The real Test Case computes reservations; the real Orchestrator decides and publishes its diagnostic.
A collection double supplies one fixed child view. Only the concurrent Suite allowance is held by
the fixture, without running a Suite. Request-entry observations are inherited from the thin child adapter.
The fault is injected by early FreeReservedEvents on a started child, not by corrupting indices or interfaces.
This tests the missing-reservation invariant; hard Event Buffer Reset mechanics are not reproduced.
Three later helper calls must retain Error without another diagnostic or unexpected dispatch.
Expected diagnostics stay in local capture. The surrounding Assertions use the normal selftest publisher.
The real subject binds only local storage; expected findings remain in that storage.
Checking Assertions retain the outer selftest publisher. Each run reinitializes the subject.
</description>
*)
{endregion}
FUNCTION_BLOCK Test_ActiveReservationLoss EXTENDS TestCaseBase
VAR
    FSubject : EventBuffer;
    FEvents : ARRAY[1..BufferLength] OF ST_Event;
    FFifo : ST_FifoStatus;
    FBufferStatus : ST_EventBufferStatus;
    FPerformed : BOOL;
    FChecked : BOOL;
    FSubjectParent : I_TestSuite;
    FChild : ReservationChildProbe;
    FOrchestrator : OrchestratorProbe;
    FCollection : OrchestrationCollectionDouble;
    FChildren : ARRAY[1..1] OF I_Orchestratable;
    FOwnerReserved : UINT;
    FStep : INT;
    FObservationCalls : UINT;
    FPrecondition : AssertTrue;
    FPreconditionMatches : BOOL;
    FFailureDetection : AssertTrue;
    FFailureDetectionMatches : BOOL;
    FStateAndCounts : AssertTrue;
    FStateAndCountsMatches : BOOL;
    FHeldError : AssertTrue;
    FHeldErrorMatches : BOOL;
    FSingleDiagnostic : AssertTrue;
    FSingleDiagnosticMatches : BOOL;
    FRequestBoundary : AssertTrue;
    FRequestBoundaryMatches : BOOL;
    FAccounting : AssertTrue;
    FAccountingMatches : BOOL;
    FCaptureIntegrity : AssertTrue;
    FCaptureIntegrityMatches : BOOL;
END_VAR
VAR CONSTANT
    ChildExecutionBudget : UINT := 11;
    ConfigureExecution : INT := 4;
    BufferLength : UINT := 65;
    ObservationCalls : UINT := 3;
    ExpectedResetRequests : UINT := 1;
    ExpectedStartRequests : UINT := 1;
    Setup : INT := 0;
    PrepareChild : INT := 1;
    TriggerFailure : INT := 2;
    ObserveFailure : INT := 3;
END_VAR

SUPER^();

{region 'Documentation'}
(*!
<summary>Contributes each checking Assertion once.</summary>
*)
{endregion}
METHOD PROTECTED AggregateResults
VAR_INPUT
    Aggregator : I_ResultAggregator; //! Borrowed result sink owned by the outer Test Case; add this test's checking Assertions without resetting or retaining the sink.
END_VAR
Aggregator.AddProvider(Provider := FPrecondition);
Aggregator.AddProvider(Provider := FFailureDetection);
Aggregator.AddProvider(Provider := FStateAndCounts);
Aggregator.AddProvider(Provider := FHeldError);
Aggregator.AddProvider(Provider := FSingleDiagnostic);
Aggregator.AddProvider(Provider := FRequestBoundary);
Aggregator.AddProvider(Provider := FAccounting);
Aggregator.AddProvider(Provider := FCaptureIntegrity);
END_METHOD

{region 'Documentation'}
(*!
<summary>Supplies only the child identity before initialization.</summary>
*)
{endregion}
METHOD PUBLIC BindSubjectParent
VAR_INPUT
    Parent : I_TestSuite; //! Borrowed identity parent retained for isolated subject initialization; keep the Suite alive through subject use.
END_VAR
FSubjectParent := Parent;
END_METHOD

{region 'Documentation'}
(*!
<summary>Calls the real helper and child and retains accounting observations.</summary>
*)
{endregion}
METHOD PRIVATE CallSubject
VAR_INPUT
    Task : E_OrchestratorTask; //! Orchestration task assigned for this controlled subject call.
END_VAR
FOrchestrator(Task := Task);
FAccountingMatches := FAccountingMatches
    AND (FSubject.ReservedEntryCount = FOwnerReserved + FChild.ReservedEntryCount);
FChild();
FCaptureIntegrityMatches := FCaptureIntegrityMatches
    AND NOT FFifo.ConfigError AND NOT FFifo.IndexError
    AND (FBufferStatus.LostEventCount = 0)
    AND NOT FCollection.InvalidAccess AND NOT FCollection.TraceOverflow;
END_METHOD

{region 'Documentation'}
(*!
<summary>Checks the single retained Orchestrator Error and exact dispatch counts.</summary>
*)
{endregion}
METHOD PRIVATE CheckDiagnostic
VAR
    Index : UINT;
    ErrorCount : UINT;
    PayloadMatches : BOOL := TRUE;
END_VAR
FOR Index := 1 TO BufferLength DO
    IF (FEvents[Index].SequenceId > 0) AND (FEvents[Index].Severity = E_EventSeverity.Error) THEN
        ErrorCount := ErrorCount + 1;
        PayloadMatches := PayloadMatches
            AND (FEvents[Index].OwnerScope = E_OwnerScope.Framework)
            AND (FEvents[Index].EventType = E_EventType.Framework)
            AND (FEvents[Index].State = E_State.Error)
            AND (FEvents[Index].Name = CONCAT(Name, '.Orchestrator'))
            AND (FEvents[Index].Message <> '');
    END_IF;
END_FOR;
FSingleDiagnosticMatches := (ErrorCount = 1) AND PayloadMatches;
FRequestBoundaryMatches := FChild.RequestsReserved
    AND (FChild.ResetRequestCount = ExpectedResetRequests)
    AND (FChild.StartRequestCount = ExpectedStartRequests);
END_METHOD

{region 'Documentation'}
(*!
<summary>Requires all checking Assertions to be initialized.</summary>
*)
{endregion}
METHOD PROTECTED CheckInitialization : BOOL //! TRUE when the inherited initialization check and this concrete fixture check both accept the setup.
CheckInitialization := FALSE;
IF NOT SUPER^.CheckInitialization() OR (FSubjectParent = 0) THEN
    RETURN;
END_IF;

CheckInitialization := FPrecondition.IsInitialized
    AND FFailureDetection.IsInitialized
    AND FStateAndCounts.IsInitialized
    AND FHeldError.IsInitialized
    AND FSingleDiagnostic.IsInitialized
    AND FRequestBoundary.IsInitialized
    AND FAccounting.IsInitialized
    AND FCaptureIntegrity.IsInitialized;
END_METHOD

{region 'Documentation'}
(*!
<summary>Initializes the checking Assertions for one test state.</summary>
*)
{endregion}
METHOD PROTECTED Configure
FPreparationStateCount := 0;
FTestStateCount := 1;
FPrecondition.Initialize(Parent := THIS^,
    AssertionName := 'Precondition');
FFailureDetection.Initialize(Parent := THIS^,
    AssertionName := 'FailureDetection');
FStateAndCounts.Initialize(Parent := THIS^,
    AssertionName := 'StateAndCounts');
FHeldError.Initialize(Parent := THIS^,
    AssertionName := 'HeldError');
FSingleDiagnostic.Initialize(Parent := THIS^,
    AssertionName := 'SingleDiagnostic');
FRequestBoundary.Initialize(Parent := THIS^,
    AssertionName := 'RequestBoundary');
FAccounting.Initialize(Parent := THIS^,
    AssertionName := 'Accounting');
FCaptureIntegrity.Initialize(Parent := THIS^,
    AssertionName := 'CaptureIntegrity');
END_METHOD

{region 'Documentation'}
(*!
<summary>Binds a real child and Orchestrator to fixed isolated storage.</summary>
*)
{endregion}
METHOD PRIVATE InitializeArrangement
VAR
    Config : ST_TestCaseConfig;
END_VAR
IF NOT FSubject.Initialize(Buffer := FEvents,
    FifoControl := FFifo,
    Status := FBufferStatus) THEN
    Error(Message := 'Reservation error capture initialization failed.');
    RETURN;
END_IF;
FOwnerReserved := 0;
FChild.BindPublisher(Publisher := FSubject);
FChild.ClearRequestTrace();
FChild.ExecutionSlot := 1;
IF NOT FChild.Initialize(Parent := FSubjectParent,
    TestName := 'LostReservationChild',
    Config := Config) THEN
    Error(Message := 'Reservation error child initialization failed.');
    RETURN;
END_IF;
FChild();
FChildren[1] := FChild;
IF NOT FCollection.Initialize(Count := 1,
    Children := FChildren) THEN
    Error(Message := 'Reservation error collection initialization failed.');
    RETURN;
END_IF;
FOrchestrator.BindPublisher(Publisher := FSubject);
IF NOT FOrchestrator.Initialize(Collection := FCollection,
    Name := Name) THEN
    Error(Message := 'Reservation error Orchestrator initialization failed.');
    RETURN;
END_IF;
IF NOT FSubject.ReserveSpace(EntryCount := GVL_Constants.TestSuiteResetEventCount,
    HeadroomEntryCount := Param_EventBuffer.EventBufferResetHeadroom,
    OwnerReservedEntryCount := FOwnerReserved) THEN
    Error(Message := 'Reservation error concurrent owner setup failed.');
    RETURN;
END_IF;
FPreconditionMatches := FPreconditionMatches AND FChild.IsInitialized
    AND FFifo.BufferEmpty AND (FSubject.Capacity = BufferLength - 1);
END_METHOD

{region 'Documentation'}
(*!
<summary>Removes setup events and replaces the fixture owner allowance; child configuration remains unchanged.</summary>
*)
{endregion}
METHOD PRIVATE PrepareExecution
VAR
    Watermark : UDINT;
END_VAR
Watermark := FBufferStatus.SequenceId;
FSubject.ProcessDeleteRequest(SequenceId := Watermark);
IF NOT FSubject.FreeReservedSpace(EntryCount := FOwnerReserved,
    OwnerReservedEntryCount := FOwnerReserved) THEN
    Error(Message := 'Could not release Reset fixture allowance.');
    RETURN;
END_IF;
IF NOT FSubject.ReserveSpace(EntryCount := GVL_Constants.TestSuiteExecutionEventCount,
    HeadroomEntryCount := Param_EventBuffer.EventBufferExecutionHeadroom,
    OwnerReservedEntryCount := FOwnerReserved) THEN
    Error(Message := 'Could not reserve execution fixture allowance.');
    RETURN;
END_IF;
FPreconditionMatches := FPreconditionMatches AND FFifo.BufferEmpty
    AND (Watermark = 0) AND (FChild.ReservedEntryCount = 0);
END_METHOD

{region 'Documentation'}
(*!
<summary>Completes abort without asynchronous work.</summary>
*)
{endregion}
METHOD PROTECTED ProcessAbort
VAR_INPUT
    Enable : BOOL; //! Phase permission supplied by the owning Test Case; FALSE does not authorize progression, while observation may continue.
END_VAR
IF Enable THEN
    CompleteAbort();
END_IF;
END_METHOD

{region 'Documentation'}
(*!
<summary>Evaluates captured observations after the scenario has finished.</summary>
*)
{endregion}
METHOD PROTECTED ProcessAssertions
VAR_INPUT
    Enable : BOOL; //! Phase permission supplied by the owning Test Case; FALSE does not authorize progression, while observation may continue.
END_VAR
VAR
    Evaluate : BOOL;
END_VAR
Evaluate := Enable AND FPerformed;
FPrecondition(Enable := Evaluate,
    State := State,
    IN := FPreconditionMatches);
FFailureDetection(Enable := Evaluate,
    State := State,
    IN := FFailureDetectionMatches);
FStateAndCounts(Enable := Evaluate,
    State := State,
    IN := FStateAndCountsMatches);
FHeldError(Enable := Evaluate,
    State := State,
    IN := FHeldErrorMatches);
FSingleDiagnostic(Enable := Evaluate,
    State := State,
    IN := FSingleDiagnosticMatches);
FRequestBoundary(Enable := Evaluate,
    State := State,
    IN := FRequestBoundaryMatches);
FAccounting(Enable := Evaluate,
    State := State,
    IN := FAccountingMatches);
FCaptureIntegrity(Enable := Evaluate,
    State := State,
    IN := FCaptureIntegrityMatches);
IF Evaluate THEN
    FChecked := TRUE;
END_IF;
END_METHOD

{region 'Documentation'}
(*!
<summary>No Preparation phase is needed.</summary>
*)
{endregion}
METHOD PROTECTED ProcessPreparations
VAR_INPUT
    // SA0033: Required override without Preparation work.
    {attribute 'analysis' := '-33'}
    Enable : BOOL; //! Phase permission supplied by the owning Test Case; FALSE does not authorize progression, while observation may continue.
END_VAR
END_METHOD

{region 'Documentation'}
(*!
<summary>Clears scenario evidence; next execution initializes a fresh local arrangement.</summary>
*)
{endregion}
METHOD PROTECTED ProcessReset
FStep := Setup;
FObservationCalls := 0;
FPerformed := FALSE;
FChecked := FALSE;
FPrecondition.Reset();
FPreconditionMatches := TRUE;
FFailureDetection.Reset();
FFailureDetectionMatches := TRUE;
FStateAndCounts.Reset();
FStateAndCountsMatches := TRUE;
FHeldError.Reset();
FHeldErrorMatches := TRUE;
FSingleDiagnostic.Reset();
FSingleDiagnosticMatches := TRUE;
FRequestBoundary.Reset();
FRequestBoundaryMatches := TRUE;
FAccounting.Reset();
FAccountingMatches := TRUE;
FCaptureIntegrity.Reset();
FCaptureIntegrityMatches := TRUE;
FSingleDiagnosticMatches := FALSE;
CompleteReset();
END_METHOD

{region 'Documentation'}
(*!
<summary>Advances one scenario phase before checking final captured observations.</summary>
*)
{endregion}
METHOD PROTECTED ProcessTests
VAR_INPUT
    Enable : BOOL; //! Phase permission supplied by the owning Test Case; FALSE does not authorize progression, while observation may continue.
END_VAR
IF NOT Enable THEN
    RETURN;
END_IF;
IF FChecked THEN
    CompleteTests();
    RETURN;
END_IF;
IF NOT FPerformed THEN
    RunScenario();
END_IF;
END_METHOD

{region 'Documentation'}
(*!
<summary>Runs one bounded scenario phase per active outer call.</summary>
*)
{endregion}
METHOD PRIVATE RunScenario
CASE FStep OF
    Setup:
        InitializeArrangement();
        FStep := PrepareChild;

    PrepareChild:
        CallSubject(Task := E_OrchestratorTask.Reset);
        IF FOrchestrator.Result = E_Result.Error THEN
            Error(Message := 'Reservation error scenario could not reset its child.');
            RETURN;
        END_IF;
        IF FOrchestrator.IsResetFinished THEN
            FPreconditionMatches := FPreconditionMatches AND FChild.IsIdle AND FChild.IsReady;
            FStep := ConfigureExecution;
        END_IF;

    ConfigureExecution:
        CallSubject(Task := E_OrchestratorTask.Idle);
        PrepareExecution();
        FStep := TriggerFailure;

    TriggerFailure:
        TriggerSubjectFailure();
        FStep := ObserveFailure;

    ObserveFailure:
        CallSubject(Task := E_OrchestratorTask.Execution);
        FFailureDetectionMatches := FFailureDetectionMatches
            AND (FOrchestrator.Result = E_Result.Error);
        FHeldErrorMatches := FHeldErrorMatches
            AND (FOrchestrator.Result = E_Result.Error)
            AND NOT FOrchestrator.IsExecutionFinished;
        FObservationCalls := FObservationCalls + 1;
        IF FObservationCalls = ObservationCalls THEN
            CheckDiagnostic();
            FAccountingMatches := FAccountingMatches
                AND (FChild.ReservedEntryCount = 0);
            IF NOT FSubject.FreeReservedSpace(EntryCount := FOwnerReserved,
                OwnerReservedEntryCount := FOwnerReserved) THEN
                Error(Message := 'Reservation error fixture cleanup failed.');
                RETURN;
            END_IF;
            FAccountingMatches := FAccountingMatches AND (FSubject.ReservedEntryCount = 0);
            FPerformed := TRUE;
        END_IF;
ELSE
    Error(Message := 'Unknown reservation error test step.');
END_CASE;
END_METHOD

{region 'Documentation'}
(*!
<summary>Releases a legitimately started child early through its public API, without changing its lifecycle.</summary>
*)
{endregion}
METHOD PRIVATE TriggerSubjectFailure
VAR
    PreviousState : E_State;
    Released : BOOL;
END_VAR
CallSubject(Task := E_OrchestratorTask.Execution);
PreviousState := FChild.State;
FPreconditionMatches := FPreconditionMatches
    AND (PreviousState >= E_State.Starting) AND (PreviousState <= E_State.Completing)
    AND (FChild.StartRequestCount = 1) AND (FChild.ReservedEntryCount = ChildExecutionBudget);
Released := FChild.FreeReservedEvents();
FStateAndCountsMatches := Released AND (FChild.State = PreviousState)
    AND (FChild.ReservedEntryCount = 0)
    AND (FSubject.ReservedEntryCount = FOwnerReserved);
END_METHOD

END_FUNCTION_BLOCK

// ---- SelfTests/TestCases/TestSuite_EventReservation/Test_HierarchicalReservationRelease.TcPOU
{region 'Documentation'}
(*!
<summary>Checks real Suite and child contributions through synchronous hierarchical release.</summary>
<description>
SuiteIntegrationSubject owns two real Test Cases with one Assertion each. Their actual
reservation methods update the same isolated EventBuffer; no child reservation markers are faked.
No lifecycle is started: release must preserve all three Uninitialized states and a retained event.
After complete execution-budget release, child Reset budgets are acquired while the Suite owns zero.
A further hierarchical release must still visit those children. Empty repeat release must be harmless.
The real subject binds only local storage; expected findings remain in that storage.
Checking Assertions retain the outer selftest publisher. Each run reinitializes the subject.
</description>
*)
{endregion}
FUNCTION_BLOCK Test_HierarchicalReservationRelease EXTENDS TestCaseBase
VAR
    FSubject : EventBuffer;
    FEvents : ARRAY[1..BufferLength] OF ST_Event;
    FFifo : ST_FifoStatus;
    FBufferStatus : ST_EventBufferStatus;
    FPerformed : BOOL;
    FChecked : BOOL;
    FSubjectParent : I_RunControl;
    FSuite : SuiteIntegrationSubject;
    FInitialization : AssertTrue;
    FInitializationMatches : BOOL;
    FExecutionContributions : AssertTrue;
    FExecutionContributionsMatches : BOOL;
    FFullRelease : AssertTrue;
    FFullReleaseMatches : BOOL;
    FRepeatedRelease : AssertTrue;
    FRepeatedReleaseMatches : BOOL;
    FZeroOwnerCleanup : AssertTrue;
    FZeroOwnerCleanupMatches : BOOL;
    FStatePreserved : AssertTrue;
    FStatePreservedMatches : BOOL;
    FEventsPreserved : AssertTrue;
    FEventsPreservedMatches : BOOL;
    FStorageIntegrity : AssertTrue;
    FStorageIntegrityMatches : BOOL;
END_VAR
VAR CONSTANT
    BufferLength : UINT := 97;
    ChildExecutionBudget : UINT := 11;
END_VAR

SUPER^();

{region 'Documentation'}
(*!
<summary>Contributes each checking Assertion once.</summary>
*)
{endregion}
METHOD PROTECTED AggregateResults
VAR_INPUT
    Aggregator : I_ResultAggregator; //! Borrowed result sink owned by the outer Test Case; add this test's checking Assertions without resetting or retaining the sink.
END_VAR
Aggregator.AddProvider(Provider := FInitialization);
Aggregator.AddProvider(Provider := FExecutionContributions);
Aggregator.AddProvider(Provider := FFullRelease);
Aggregator.AddProvider(Provider := FRepeatedRelease);
Aggregator.AddProvider(Provider := FZeroOwnerCleanup);
Aggregator.AddProvider(Provider := FStatePreserved);
Aggregator.AddProvider(Provider := FEventsPreserved);
Aggregator.AddProvider(Provider := FStorageIntegrity);
END_METHOD

{region 'Documentation'}
(*!
<summary>Supplies root identity only; the root never calls this isolated Suite.</summary>
*)
{endregion}
METHOD PUBLIC BindSubjectParent
VAR_INPUT
    Parent : I_RunControl; //! Borrowed identity parent retained for isolated subject initialization; keep the Run-Control alive through subject use.
END_VAR
FSubjectParent := Parent;
END_METHOD

{region 'Documentation'}
(*!
<summary>Requires all checking Assertions to be initialized.</summary>
*)
{endregion}
METHOD PROTECTED CheckInitialization : BOOL //! TRUE when the inherited initialization check and this concrete fixture check both accept the setup.
CheckInitialization := FALSE;
IF NOT SUPER^.CheckInitialization() OR (FSubjectParent = 0) THEN
    RETURN;
END_IF;

CheckInitialization := FInitialization.IsInitialized
    AND FExecutionContributions.IsInitialized
    AND FFullRelease.IsInitialized
    AND FRepeatedRelease.IsInitialized
    AND FZeroOwnerCleanup.IsInitialized
    AND FStatePreserved.IsInitialized
    AND FEventsPreserved.IsInitialized
    AND FStorageIntegrity.IsInitialized;
END_METHOD

{region 'Documentation'}
(*!
<summary>Initializes the checking Assertions for one test state.</summary>
*)
{endregion}
METHOD PROTECTED Configure
FPreparationStateCount := 0;
FTestStateCount := 1;
FInitialization.Initialize(Parent := THIS^,
    AssertionName := 'Initialization');
FExecutionContributions.Initialize(Parent := THIS^,
    AssertionName := 'ExecutionContributions');
FFullRelease.Initialize(Parent := THIS^,
    AssertionName := 'FullRelease');
FRepeatedRelease.Initialize(Parent := THIS^,
    AssertionName := 'RepeatedRelease');
FZeroOwnerCleanup.Initialize(Parent := THIS^,
    AssertionName := 'ZeroOwnerCleanup');
FStatePreserved.Initialize(Parent := THIS^,
    AssertionName := 'StatePreserved');
FEventsPreserved.Initialize(Parent := THIS^,
    AssertionName := 'EventsPreserved');
FStorageIntegrity.Initialize(Parent := THIS^,
    AssertionName := 'StorageIntegrity');
END_METHOD

{region 'Documentation'}
(*!
<summary>Checks actual subtree accounting without dispatching lifecycle requests.</summary>
*)
{endregion}
METHOD PRIVATE ExerciseBuffer
VAR
    Config : ST_TestSuiteConfig;
    FirstChild : I_TestCase;
    SecondChild : I_TestCase;
    Initialized : BOOL;
    Released : BOOL;
    SuiteReservation : E_EventReservationResult;
    FirstReservation : E_EventReservationResult;
    SecondReservation : E_EventReservationResult;
    RetainedSequence : UDINT;
END_VAR
Initialized := FSubject.Initialize(Buffer := FEvents,
    FifoControl := FFifo,
    Status := FBufferStatus);
IF NOT Initialized THEN
    Error(Message := 'Hierarchical release capture initialization failed.');
    RETURN;
END_IF;
FSuite.BindPublisher(Publisher := FSubject);
IF NOT FSuite.Initialize(Parent := FSubjectParent,
    SuiteName := 'ReservationRelease',
    Config := Config) THEN
    Error(Message := 'Hierarchical release Suite initialization failed.');
    RETURN;
END_IF;
FSuite();
FirstChild := FSuite.GetTestCase(Index := FSuite.ChildArrayLowerBound);
SecondChild := FSuite.GetTestCase(Index := FSuite.ChildArrayLowerBound + 1);
FInitializationMatches := FSuite.IsInitialized AND FirstChild.IsInitialized AND SecondChild.IsInitialized
    AND (FSuite.ChildCount = 2) AND FSuite.ChildCallsMatch;
IF FSubject.PublishEvent(Event := CreateFrameworkEvent(Name := Name,
    State := E_State.Uninitialized,
    Severity := E_EventSeverity.Info,
    Message := 'Retained across hierarchical reservation release.')) <= 0 THEN
    Error(Message := 'Hierarchical release retained event setup failed.');
    RETURN;
END_IF;
RetainedSequence := FBufferStatus.SequenceId;

SuiteReservation := FSuite.ReserveExecutionEvents();
FirstReservation := FirstChild.ReserveExecutionEvents();
SecondReservation := SecondChild.ReserveExecutionEvents();
FExecutionContributionsMatches := (SuiteReservation = E_EventReservationResult.Accepted)
    AND (FirstReservation = E_EventReservationResult.Accepted)
    AND (SecondReservation = E_EventReservationResult.Accepted)
    AND (FSuite.ReservedEntryCount = GVL_Constants.TestSuiteExecutionEventCount)
    AND (FirstChild.ReservedEntryCount = ChildExecutionBudget)
    AND (SecondChild.ReservedEntryCount = ChildExecutionBudget)
    AND (FSubject.ReservedEntryCount = GVL_Constants.TestSuiteExecutionEventCount + 2 * ChildExecutionBudget);

Released := FSuite.FreeReservedEvents();
FFullReleaseMatches := Released AND (FSuite.ReservedEntryCount = 0)
    AND (FirstChild.ReservedEntryCount = 0) AND (SecondChild.ReservedEntryCount = 0)
    AND (FSubject.ReservedEntryCount = 0);
Released := FSuite.FreeReservedEvents();
FRepeatedReleaseMatches := Released AND (FSubject.ReservedEntryCount = 0)
    AND (FSuite.ReservedEntryCount = 0)
    AND (FirstChild.ReservedEntryCount = 0) AND (SecondChild.ReservedEntryCount = 0);

FirstReservation := FirstChild.ReserveResetEvents();
SecondReservation := SecondChild.ReserveResetEvents();
FZeroOwnerCleanupMatches := (FirstReservation = E_EventReservationResult.Accepted)
    AND (SecondReservation = E_EventReservationResult.Accepted)
    AND (FSuite.ReservedEntryCount = 0)
    AND (FSubject.ReservedEntryCount = 2 * GVL_Constants.TestCaseResetEventCount);
Released := FSuite.FreeReservedEvents();
FZeroOwnerCleanupMatches := FZeroOwnerCleanupMatches AND Released
    AND (FirstChild.ReservedEntryCount = 0) AND (SecondChild.ReservedEntryCount = 0)
    AND (FSuite.ReservedEntryCount = 0) AND (FSubject.ReservedEntryCount = 0);
FStatePreservedMatches := (FSuite.State = E_State.Uninitialized)
    AND (FirstChild.State = E_State.Uninitialized) AND (SecondChild.State = E_State.Uninitialized);
FEventsPreservedMatches := (FBufferStatus.SequenceId = RetainedSequence)
    AND (FBufferStatus.DeletedSequenceId = 0) AND (FFifo.ElementCount = 1)
    AND (FEvents[FFifo.IndexOut].SequenceId = RetainedSequence);
FStorageIntegrityMatches := NOT FFifo.ConfigError AND NOT FFifo.IndexError
    AND (FBufferStatus.LostEventCount = 0);
END_METHOD

{region 'Documentation'}
(*!
<summary>Completes abort without asynchronous work.</summary>
*)
{endregion}
METHOD PROTECTED ProcessAbort
VAR_INPUT
    Enable : BOOL; //! Phase permission supplied by the owning Test Case; FALSE does not authorize progression, while observation may continue.
END_VAR
IF Enable THEN
    CompleteAbort();
END_IF;
END_METHOD

{region 'Documentation'}
(*!
<summary>Evaluates captured observations after the scenario has finished.</summary>
*)
{endregion}
METHOD PROTECTED ProcessAssertions
VAR_INPUT
    Enable : BOOL; //! Phase permission supplied by the owning Test Case; FALSE does not authorize progression, while observation may continue.
END_VAR
VAR
    Evaluate : BOOL;
END_VAR
Evaluate := Enable AND FPerformed;
FInitialization(Enable := Evaluate,
    State := State,
    IN := FInitializationMatches);
FExecutionContributions(Enable := Evaluate,
    State := State,
    IN := FExecutionContributionsMatches);
FFullRelease(Enable := Evaluate,
    State := State,
    IN := FFullReleaseMatches);
FRepeatedRelease(Enable := Evaluate,
    State := State,
    IN := FRepeatedReleaseMatches);
FZeroOwnerCleanup(Enable := Evaluate,
    State := State,
    IN := FZeroOwnerCleanupMatches);
FStatePreserved(Enable := Evaluate,
    State := State,
    IN := FStatePreservedMatches);
FEventsPreserved(Enable := Evaluate,
    State := State,
    IN := FEventsPreservedMatches);
FStorageIntegrity(Enable := Evaluate,
    State := State,
    IN := FStorageIntegrityMatches);
IF Evaluate THEN
    FChecked := TRUE;
END_IF;
END_METHOD

{region 'Documentation'}
(*!
<summary>No Preparation phase is needed.</summary>
*)
{endregion}
METHOD PROTECTED ProcessPreparations
VAR_INPUT
    // SA0033: Required override without Preparation work.
    {attribute 'analysis' := '-33'}
    Enable : BOOL; //! Phase permission supplied by the owning Test Case; FALSE does not authorize progression, while observation may continue.
END_VAR
END_METHOD

{region 'Documentation'}
(*!
<summary>Resets observations and schedules a fresh subject initialization.</summary>
*)
{endregion}
METHOD PROTECTED ProcessReset
FPerformed := FALSE;
FChecked := FALSE;
FInitialization.Reset();
FInitializationMatches := FALSE;
FExecutionContributions.Reset();
FExecutionContributionsMatches := FALSE;
FFullRelease.Reset();
FFullReleaseMatches := FALSE;
FRepeatedRelease.Reset();
FRepeatedReleaseMatches := FALSE;
FZeroOwnerCleanup.Reset();
FZeroOwnerCleanupMatches := FALSE;
FStatePreserved.Reset();
FStatePreservedMatches := FALSE;
FEventsPreserved.Reset();
FEventsPreservedMatches := FALSE;
FStorageIntegrity.Reset();
FStorageIntegrityMatches := FALSE;
CompleteReset();
END_METHOD

{region 'Documentation'}
(*!
<summary>Runs the bounded scenario once before Assertion evaluation.</summary>
*)
{endregion}
METHOD PROTECTED ProcessTests
VAR_INPUT
    Enable : BOOL; //! Phase permission supplied by the owning Test Case; FALSE does not authorize progression, while observation may continue.
END_VAR
IF NOT Enable THEN
    RETURN;
END_IF;
IF FChecked THEN
    CompleteTests();
    RETURN;
END_IF;

IF NOT FPerformed THEN
    ExerciseBuffer();
    FPerformed := TRUE;
END_IF;
END_METHOD

END_FUNCTION_BLOCK

// ---- SelfTests/TestCases/TestSuite_EventReservation/Test_LateResetReservationRelease.TcPOU
{region 'Documentation'}
(*!
<summary>Checks hierarchical early release after a real Suite Reset timeout while children still reset.</summary>
<description>

Controlled concrete Reset work

The Suite and Orchestrator are real. Both real children remain in their concrete Reset hook
until the scenario releases it; their normal five-second deadlines remain active.
The Suite uses a 100 ms Reset timeout. No timer/state field is manipulated and no duration is benchmarked.

Accepted failure-path gap

After the Suite reaches Completed/Error, the test performs parent-owned hierarchical release.
Three further calls must retain resetting children with zero reservations and no new dispatch.
The hooks are then released: children publish late Idle transitions while the Suite's final result
and finalization remain unchanged. This deliberately checks the accepted temporary coverage gap,
not a general guarantee for arbitrarily many events after faulty early release.
The real subject binds only local storage; expected findings remain in that storage.
Checking Assertions retain the outer selftest publisher. Each run reinitializes the subject.
</description>
*)
{endregion}
FUNCTION_BLOCK Test_LateResetReservationRelease EXTENDS TestCaseBase
VAR
    FSubject : EventBuffer;
    FEvents : ARRAY[1..BufferLength] OF ST_Event;
    FFifo : ST_FifoStatus;
    FBufferStatus : ST_EventBufferStatus;
    FPerformed : BOOL;
    FChecked : BOOL;
    FSubjectParent : I_RunControl;
    FSuite : ReservationSuiteProbe;
    FFirstChild : I_TestCase;
    FSecondChild : I_TestCase;
    FStep : INT;
    FHoldCalls : UINT;
    FReleaseSequence : UDINT;
    FResetAdmission : AssertTrue;
    FResetAdmissionMatches : BOOL;
    FOwnerFinalization : AssertTrue;
    FOwnerFinalizationMatches : BOOL;
    FEarlyRelease : AssertTrue;
    FEarlyReleaseMatches : BOOL;
    FRepeatedRelease : AssertTrue;
    FRepeatedReleaseMatches : BOOL;
    FLateCompletion : AssertTrue;
    FLateCompletionMatches : BOOL;
    FStableOwner : AssertTrue;
    FStableOwnerMatches : BOOL;
    FAccounting : AssertTrue;
    FAccountingMatches : BOOL;
    FEventEvidence : AssertTrue;
    FEventEvidenceMatches : BOOL;
END_VAR
VAR CONSTANT
    BufferLength : UINT := 97;
    HoldCalls : UINT := 3;
    Setup : INT := 0;
    WaitForOwnerCompletion : INT := 1;
    ObserveReleasedChildren : INT := 2;
    WaitForChildCompletion : INT := 3;
END_VAR

SUPER^();

{region 'Documentation'}
(*!
<summary>Contributes each checking Assertion once.</summary>
*)
{endregion}
METHOD PROTECTED AggregateResults
VAR_INPUT
    Aggregator : I_ResultAggregator; //! Borrowed result sink owned by the outer Test Case; add this test's checking Assertions without resetting or retaining the sink.
END_VAR
Aggregator.AddProvider(Provider := FResetAdmission);
Aggregator.AddProvider(Provider := FOwnerFinalization);
Aggregator.AddProvider(Provider := FEarlyRelease);
Aggregator.AddProvider(Provider := FRepeatedRelease);
Aggregator.AddProvider(Provider := FLateCompletion);
Aggregator.AddProvider(Provider := FStableOwner);
Aggregator.AddProvider(Provider := FAccounting);
Aggregator.AddProvider(Provider := FEventEvidence);
END_METHOD

{region 'Documentation'}
(*!
<summary>Supplies root identity only; the outer root does not execute the isolated Suite.</summary>
*)
{endregion}
METHOD PUBLIC BindSubjectParent
VAR_INPUT
    Parent : I_RunControl; //! Borrowed identity parent retained for isolated subject initialization; keep the Run-Control alive through subject use.
END_VAR
FSubjectParent := Parent;
END_METHOD

{region 'Documentation'}
(*!
<summary>Compares real local contributions with the buffer aggregate and checks continuous child calls.</summary>
*)
{endregion}
METHOD PRIVATE CheckAccounting
FAccountingMatches := FAccountingMatches
    AND (FSubject.ReservedEntryCount = FSuite.ReservedEntryCount
        + FFirstChild.ReservedEntryCount + FSecondChild.ReservedEntryCount)
    AND FSuite.ChildCallsMatch
    AND NOT FFifo.ConfigError AND NOT FFifo.IndexError
    AND (FBufferStatus.LostEventCount = 0);
END_METHOD

{region 'Documentation'}
(*!
<summary>Checks one parent finalization and child Idle events after release, without promising late-event reservation coverage.</summary>
*)
{endregion}
METHOD PRIVATE CheckFinalEvents
VAR
    Index : UINT;
    SuiteResults : UINT;
    SuiteAggregations : UINT;
    SuiteCompletions : UINT;
    FirstLateIdle : UINT;
    SecondLateIdle : UINT;
    PayloadMatches : BOOL := TRUE;
END_VAR
FOR Index := 1 TO BufferLength DO
    IF FEvents[Index].SequenceId = 0 THEN
        CONTINUE;
    END_IF;
    IF FEvents[Index].EventType = E_EventType.StateTransition THEN
        PayloadMatches := PayloadMatches
            AND (FEvents[Index].State <> E_State.Aborting)
            AND (FEvents[Index].State <> E_State.AbortingFromError);
    END_IF;
    IF FEvents[Index].Name = FSuite.Name THEN
        CASE FEvents[Index].EventType OF
            E_EventType.Result:
                SuiteResults := SuiteResults + 1;
                PayloadMatches := PayloadMatches AND (FEvents[Index].Result = E_Result.Error);
            E_EventType.Aggregation:
                SuiteAggregations := SuiteAggregations + 1;
            E_EventType.StateTransition:
                IF FEvents[Index].State = E_State.Completed THEN
                    SuiteCompletions := SuiteCompletions + 1;
                    PayloadMatches := PayloadMatches AND (FEvents[Index].SequenceId <= FReleaseSequence);
                END_IF;
        END_CASE;
    ELSIF (FEvents[Index].SequenceId > FReleaseSequence)
        AND (FEvents[Index].EventType = E_EventType.StateTransition)
        AND (FEvents[Index].State = E_State.Idle) THEN
        IF FEvents[Index].Name = FFirstChild.Name THEN
            FirstLateIdle := FirstLateIdle + 1;
        ELSIF FEvents[Index].Name = FSecondChild.Name THEN
            SecondLateIdle := SecondLateIdle + 1;
        END_IF;
    END_IF;
END_FOR;
FEventEvidenceMatches := PayloadMatches
    AND (SuiteResults = 1) AND (SuiteAggregations = 1) AND (SuiteCompletions = 1)
    AND (FirstLateIdle = 1) AND (SecondLateIdle = 1);
END_METHOD

{region 'Documentation'}
(*!
<summary>Requires all checking Assertions to be initialized.</summary>
*)
{endregion}
METHOD PROTECTED CheckInitialization : BOOL //! TRUE when the inherited initialization check and this concrete fixture check both accept the setup.
CheckInitialization := FALSE;
IF NOT SUPER^.CheckInitialization() OR (FSubjectParent = 0) THEN
    RETURN;
END_IF;

CheckInitialization := FResetAdmission.IsInitialized
    AND FOwnerFinalization.IsInitialized
    AND FEarlyRelease.IsInitialized
    AND FRepeatedRelease.IsInitialized
    AND FLateCompletion.IsInitialized
    AND FStableOwner.IsInitialized
    AND FAccounting.IsInitialized
    AND FEventEvidence.IsInitialized;
END_METHOD

{region 'Documentation'}
(*!
<summary>Initializes the checking Assertions for one test state.</summary>
*)
{endregion}
METHOD PROTECTED Configure
FPreparationStateCount := 0;
FTestStateCount := 1;
FResetAdmission.Initialize(Parent := THIS^,
    AssertionName := 'ResetAdmission');
FOwnerFinalization.Initialize(Parent := THIS^,
    AssertionName := 'OwnerFinalization');
FEarlyRelease.Initialize(Parent := THIS^,
    AssertionName := 'EarlyRelease');
FRepeatedRelease.Initialize(Parent := THIS^,
    AssertionName := 'RepeatedRelease');
FLateCompletion.Initialize(Parent := THIS^,
    AssertionName := 'LateCompletion');
FStableOwner.Initialize(Parent := THIS^,
    AssertionName := 'StableOwner');
FAccounting.Initialize(Parent := THIS^,
    AssertionName := 'Accounting');
FEventEvidence.Initialize(Parent := THIS^,
    AssertionName := 'EventEvidence');
END_METHOD

{region 'Documentation'}
(*!
<summary>Binds the real hierarchy and requests Reset with a shorter Suite deadline than its children.</summary>
*)
{endregion}
METHOD PRIVATE InitializeArrangement
VAR
    Config : ST_TestSuiteConfig;
END_VAR
IF NOT FSubject.Initialize(Buffer := FEvents,
    FifoControl := FFifo,
    Status := FBufferStatus) THEN
    Error(Message := 'Late Reset capture initialization failed.');
    RETURN;
END_IF;
FSuite.BindPublisher(Publisher := FSubject,
    AllowResetCompletion := FALSE);
Config.ResetTimeout := T#100ms;
IF NOT FSuite.Initialize(Parent := FSubjectParent,
    SuiteName := 'LateResetRelease',
    Config := Config) THEN
    Error(Message := 'Late Reset Suite initialization failed.');
    RETURN;
END_IF;
FFirstChild := FSuite.GetTestCase(Index := FSuite.ChildArrayLowerBound);
FSecondChild := FSuite.GetTestCase(Index := FSuite.ChildArrayLowerBound + 1);
IF FSuite.ReserveResetEvents() <> E_EventReservationResult.Accepted THEN
    Error(Message := 'Late Reset Suite reservation failed.');
    RETURN;
END_IF;
FSuite.RequestReset();
END_METHOD

{region 'Documentation'}
(*!
<summary>Completes abort without asynchronous work.</summary>
*)
{endregion}
METHOD PROTECTED ProcessAbort
VAR_INPUT
    Enable : BOOL; //! Phase permission supplied by the owning Test Case; FALSE does not authorize progression, while observation may continue.
END_VAR
IF Enable THEN
    CompleteAbort();
END_IF;
END_METHOD

{region 'Documentation'}
(*!
<summary>Evaluates captured observations after the scenario has finished.</summary>
*)
{endregion}
METHOD PROTECTED ProcessAssertions
VAR_INPUT
    Enable : BOOL; //! Phase permission supplied by the owning Test Case; FALSE does not authorize progression, while observation may continue.
END_VAR
VAR
    Evaluate : BOOL;
END_VAR
Evaluate := Enable AND FPerformed;
FResetAdmission(Enable := Evaluate,
    State := State,
    IN := FResetAdmissionMatches);
FOwnerFinalization(Enable := Evaluate,
    State := State,
    IN := FOwnerFinalizationMatches);
FEarlyRelease(Enable := Evaluate,
    State := State,
    IN := FEarlyReleaseMatches);
FRepeatedRelease(Enable := Evaluate,
    State := State,
    IN := FRepeatedReleaseMatches);
FLateCompletion(Enable := Evaluate,
    State := State,
    IN := FLateCompletionMatches);
FStableOwner(Enable := Evaluate,
    State := State,
    IN := FStableOwnerMatches);
FAccounting(Enable := Evaluate,
    State := State,
    IN := FAccountingMatches);
FEventEvidence(Enable := Evaluate,
    State := State,
    IN := FEventEvidenceMatches);
IF Evaluate THEN
    FChecked := TRUE;
END_IF;
END_METHOD

{region 'Documentation'}
(*!
<summary>No Preparation phase is needed.</summary>
*)
{endregion}
METHOD PROTECTED ProcessPreparations
VAR_INPUT
    // SA0033: Required override without Preparation work.
    {attribute 'analysis' := '-33'}
    Enable : BOOL; //! Phase permission supplied by the owning Test Case; FALSE does not authorize progression, while observation may continue.
END_VAR
END_METHOD

{region 'Documentation'}
(*!
<summary>Clears observations; next execution initializes fresh isolated storage and hierarchy.</summary>
*)
{endregion}
METHOD PROTECTED ProcessReset
FStep := Setup;
FHoldCalls := 0;
FReleaseSequence := 0;
FPerformed := FALSE;
FChecked := FALSE;
FResetAdmission.Reset();
FResetAdmissionMatches := TRUE;
FOwnerFinalization.Reset();
FOwnerFinalizationMatches := TRUE;
FEarlyRelease.Reset();
FEarlyReleaseMatches := TRUE;
FRepeatedRelease.Reset();
FRepeatedReleaseMatches := TRUE;
FLateCompletion.Reset();
FLateCompletionMatches := TRUE;
FStableOwner.Reset();
FStableOwnerMatches := TRUE;
FAccounting.Reset();
FAccountingMatches := TRUE;
FEventEvidence.Reset();
FEventEvidenceMatches := TRUE;
FEventEvidenceMatches := FALSE;
CompleteReset();
END_METHOD

{region 'Documentation'}
(*!
<summary>Calls the isolated hierarchy at most once per active cycle; outer timeout bounds non-completion.</summary>
*)
{endregion}
METHOD PROTECTED ProcessTests
VAR_INPUT
    Enable : BOOL; //! Phase permission supplied by the owning Test Case; FALSE does not authorize progression, while observation may continue.
END_VAR
IF NOT Enable THEN
    RETURN;
END_IF;
IF FChecked THEN
    CompleteTests();
    RETURN;
END_IF;
IF NOT FPerformed THEN
    RunScenario();
END_IF;
END_METHOD

{region 'Documentation'}
(*!
<summary>Releases the completed parent and still-resetting children without changing their states.</summary>
*)
{endregion}
METHOD PRIVATE ReleaseSubtree
VAR
    Released : BOOL;
END_VAR
FReleaseSequence := FBufferStatus.SequenceId;
Released := FSuite.FreeReservedEvents();
FEarlyReleaseMatches := Released
    AND (FSuite.State = E_State.Completed)
    AND (FFirstChild.State = E_State.Reset) AND (FSecondChild.State = E_State.Reset)
    AND (FSuite.ReservedEntryCount = 0)
    AND (FFirstChild.ReservedEntryCount = 0) AND (FSecondChild.ReservedEntryCount = 0)
    AND (FSubject.ReservedEntryCount = 0)
    AND (FBufferStatus.SequenceId = FReleaseSequence);
Released := FSuite.FreeReservedEvents();
FRepeatedReleaseMatches := Released AND (FSubject.ReservedEntryCount = 0)
    AND (FBufferStatus.SequenceId = FReleaseSequence);
END_METHOD

{region 'Documentation'}
(*!
<summary>Advances one explicit failure-path checkpoint per task call.</summary>
*)
{endregion}
METHOD PRIVATE RunScenario
CASE FStep OF
    Setup:
        InitializeArrangement();
        FStep := WaitForOwnerCompletion;

    WaitForOwnerCompletion:
        FSuite();
        CheckAccounting();
        IF FSuite.IsComplete THEN
            FOwnerFinalizationMatches := (FSuite.Result = E_Result.Error)
                AND FSuite.HasResetTimeout
                AND (FFirstChild.State = E_State.Reset)
                AND (FSecondChild.State = E_State.Reset)
                AND FSuite.ResetRequestsMatch;
            FResetAdmissionMatches := (FSuite.ReservedEntryCount = GVL_Constants.TestSuiteResetEventCount)
                AND (FFirstChild.ReservedEntryCount = GVL_Constants.TestCaseResetEventCount)
                AND (FSecondChild.ReservedEntryCount = GVL_Constants.TestCaseResetEventCount);
            ReleaseSubtree();
            FStep := ObserveReleasedChildren;
        END_IF;

    ObserveReleasedChildren:
        FSuite();
        CheckAccounting();
        FStableOwnerMatches := FStableOwnerMatches AND FSuite.IsComplete
            AND (FSuite.Result = E_Result.Error) AND FSuite.ResetRequestsMatch;
        FEarlyReleaseMatches := FEarlyReleaseMatches
            AND (FFirstChild.State = E_State.Reset) AND (FSecondChild.State = E_State.Reset)
            AND (FSubject.ReservedEntryCount = 0)
            AND (FBufferStatus.SequenceId = FReleaseSequence);
        FHoldCalls := FHoldCalls + 1;
        IF FHoldCalls = HoldCalls THEN
            FSuite.AllowChildResetCompletion();
            FStep := WaitForChildCompletion;
        END_IF;

    WaitForChildCompletion:
        FSuite();
        CheckAccounting();
        FStableOwnerMatches := FStableOwnerMatches AND FSuite.IsComplete
            AND (FSuite.Result = E_Result.Error) AND FSuite.ResetRequestsMatch;
        IF (FFirstChild.State = E_State.Idle) AND FFirstChild.IsReady
            AND (FSecondChild.State = E_State.Idle) AND FSecondChild.IsReady THEN
            FLateCompletionMatches := (FSubject.ReservedEntryCount = 0)
                AND (FBufferStatus.SequenceId > FReleaseSequence)
                AND FSuite.ChildCallsMatch;
            CheckFinalEvents();
            IF NOT FSuite.FreeReservedEvents() THEN
                Error(Message := 'Final repeated subtree release failed.');
                RETURN;
            END_IF;
            FRepeatedReleaseMatches := FRepeatedReleaseMatches AND (FSubject.ReservedEntryCount = 0);
            FPerformed := TRUE;
        END_IF;
ELSE
    Error(Message := 'Unknown late Reset release test step.');
END_CASE;
END_METHOD

END_FUNCTION_BLOCK

// ---- SelfTests/TestCases/TestSuite_EventReservation/Helper/ReservationSuiteProbe.TcPOU
{region 'Documentation'}
(*!
<summary>Composes two real children with a controllable concrete Reset completion.</summary>
<description>
Production TestSuiteBase and Orchestrator own all lifecycle, scheduling and reservation decisions.
BindPublisher assigns every dependency before initialization; AllowResetCompletion can hold both
children in their ordinary Reset hooks. AllowChildResetCompletion releases those hooks later.
No state, timer or reservation field is changed by the adapter. Children keep a five-second Reset
timeout while the test chooses a shorter Suite timeout. Request counters expose redispatch.
</description>
*)
{endregion}
FUNCTION_BLOCK ReservationSuiteProbe EXTENDS TestSuiteBase
VAR
    FFirst : ReservationResetChild;
    FSecond : ReservationResetChild;
    FTestCases : ARRAY[4..6] OF I_TestCase;
    FRealOrchestrator : OrchestratorProbe;
    FAllowResetCompletion : BOOL := TRUE;
    FBodyCallCount : UDINT;
    FConfigureCount : UINT;
END_VAR

FBodyCallCount := FBodyCallCount + 1;
SUPER^();

{region 'Documentation'}
(*!
<summary>Lets subsequent child calls complete their concrete Reset hooks.</summary>
*)
{endregion}
METHOD PUBLIC AllowChildResetCompletion
FAllowResetCompletion := TRUE;
END_METHOD

{region 'Documentation'}
(*!
<summary>Binds every producer before Initialize; never modifies the global publisher.</summary>
*)
{endregion}
METHOD PUBLIC BindPublisher
VAR_INPUT
    Publisher : I_EventPublisher; //! Nonzero isolated event publisher retained before subject initialization; keep it alive through all subject use.
    AllowResetCompletion : BOOL := TRUE; //! Reset-completion permission propagated to the controlled children.
END_VAR
FAllowResetCompletion := AllowResetCompletion;
FEventPublisher := Publisher;
FRealOrchestrator.BindPublisher(Publisher := Publisher);
FOrchestrator := FRealOrchestrator;
FFirst.BindPublisher(Publisher := Publisher);
FSecond.BindPublisher(Publisher := Publisher);
FFirst.ClearRequestTrace();
FSecond.ClearRequestTrace();
FBodyCallCount := 0;
FConfigureCount := 0;
END_METHOD

{region 'Documentation'}
(*!
<summary>Confirms one concrete child call per Suite call, including Reset and Completed.</summary>
*)
{endregion}
{attribute 'monitoring' := 'call'}
PROPERTY PUBLIC ChildCallsMatch : BOOL //! Confirms one concrete child call per Suite call, including Reset and Completed.
GET
ChildCallsMatch := (FFirst.BodyCallCount = FBodyCallCount) AND (FSecond.BodyCallCount = FBodyCallCount);
END_GET
END_PROPERTY

{region 'Documentation'}
(*!
<summary>Initializes and registers two real children serially in a shifted array with one unused slot.</summary>
*)
{endregion}
METHOD PROTECTED Configure
VAR_IN_OUT
    // SA0167: Borrowed setup builder; no temporary instance is created.
    {attribute 'analysis' := '-167'}
    Builder : TestSuiteConfigurationBuilder; //! Borrowed owner configuration builder used only during this Configure call; register this owner's concrete children.
END_VAR
VAR
    Config : ST_TestCaseConfig;
END_VAR
FConfigureCount := FConfigureCount + 1;
Builder.Initialize(Mode := E_OrchestrationMode.Serial,
    TestCases := FTestCases);
Config.ResetTimeout := T#5s;
FFirst.Initialize(Parent := THIS^,
    TestName := 'First',
    Config := Config);
FSecond.Initialize(Parent := THIS^,
    TestName := 'Second',
    Config := Config);
Builder.Register(TestCase := FFirst);
Builder.Register(TestCase := FSecond);
END_METHOD

{region 'Documentation'}
(*!
<summary>Distinguishes Reset/repeat from reinitializing the subject.</summary>
*)
{endregion}
{attribute 'monitoring' := 'call'}
PROPERTY PUBLIC ConfigureCount : UINT //! Distinguishes Reset/repeat from reinitializing the subject.
GET
ConfigureCount := FConfigureCount;
END_GET
END_PROPERTY

{region 'Documentation'}
(*!
<summary>Resolves the actual registered array index without executing the child.</summary>
*)
{endregion}
METHOD PUBLIC GetTestCase : I_TestCase //! Typed child interface at the original array index; zero when no entry is available.
VAR_INPUT
    Index : DINT; //! Original occupied child-array index, rather than an ordinal position.
END_VAR
GetTestCase := 0;
IF (ChildCount = 0) OR (Index < ChildArrayLowerBound)
    OR (DINT_TO_LINT(Index) >= DINT_TO_LINT(ChildArrayLowerBound) + UINT_TO_LINT(ChildCount)) THEN
    RETURN;
END_IF;
GetTestCase := FTestCases[Index];
END_METHOD

{region 'Documentation'}
(*!
<summary>Calls both children once per initialized Suite call; the helper requests their lifecycle actions.</summary>
*)
{endregion}
METHOD PROTECTED ProcessTestCases
FFirst(AllowResetCompletion := FAllowResetCompletion);
FSecond(AllowResetCompletion := FAllowResetCompletion);
END_METHOD

{region 'Documentation'}
(*!
<summary>Each child received exactly one Reset and no Start in the timeout scenario.</summary>
*)
{endregion}
{attribute 'monitoring' := 'call'}
PROPERTY PUBLIC ResetRequestsMatch : BOOL //! Each child received exactly one Reset and no Start in the timeout scenario.
GET
ResetRequestsMatch := (FFirst.ResetRequestCount = 1) AND (FSecond.ResetRequestCount = 1)
    AND (FFirst.StartRequestCount = 0) AND (FSecond.StartRequestCount = 0)
    AND FFirst.RequestsReserved AND FSecond.RequestsReserved;
END_GET
END_PROPERTY

END_FUNCTION_BLOCK

// ---- SelfTests/TestCases/TestSuite_EventReservation/Helper/ReservationResetChild.TcPOU
{region 'Documentation'}
(*!
<summary>Delays only the concrete Reset completion; all lifecycle and reservation processing remains inherited.</summary>
*)
{endregion}
FUNCTION_BLOCK ReservationResetChild EXTENDS ReservationChildProbe
VAR_INPUT
    AllowResetCompletion : BOOL := TRUE; //! FALSE holds the real child in Reset; TRUE permits inherited Reset completion.
END_VAR

SUPER^();

{region 'Documentation'}
(*!
<summary>Completes the concrete Reset only when released by the local scenario.</summary>
*)
{endregion}
METHOD PROTECTED ProcessReset
IF AllowResetCompletion THEN
    SUPER^.ProcessReset();
END_IF;
END_METHOD

END_FUNCTION_BLOCK

// ---- SelfTests/TestSuites/TestSuite_EventBufferReset.TcPOU
{region 'Documentation'}
(*!
<summary>Checks coordinated hard buffer reset on isolated real storage and hierarchy.</summary>
*)
{endregion}
FUNCTION_BLOCK TestSuite_EventBufferReset EXTENDS TestSuiteBase
VAR
    FEpochs : Test_BufferResetEpochs;
    FCommands : Test_BufferResetCommands;
    FActiveRun : Test_BufferResetActiveRun;
    FTestCases : ARRAY[1..TestCaseCapacity] OF I_TestCase;
END_VAR
VAR CONSTANT
    TestCaseCapacity : UINT := 3;
END_VAR

SUPER^();

{region 'Documentation'}
(*!
<summary>Initializes and registers the isolated event scenarios for serial execution.</summary>
*)
{endregion}
METHOD PROTECTED Configure
VAR_IN_OUT
    // SA0167: Borrowed owner builder; no temporary instance is created.
    {attribute 'analysis' := '-167'}
    Builder : TestSuiteConfigurationBuilder; //! Borrowed owner configuration builder used only during this Configure call; register this owner's concrete children.
END_VAR
VAR
    TestConfig : ST_TestCaseConfig;
END_VAR
Builder.Initialize(Mode := E_OrchestrationMode.Serial,
    TestCases := FTestCases);
FEpochs.Initialize(Parent := THIS^,
    TestName := 'Epochs',
    Config := TestConfig);
Builder.Register(TestCase := FEpochs);
FCommands.Initialize(Parent := THIS^,
    TestName := 'Commands',
    Config := TestConfig);
Builder.Register(TestCase := FCommands);
FActiveRun.Initialize(Parent := THIS^,
    TestName := 'ActiveRun',
    Config := TestConfig);
Builder.Register(TestCase := FActiveRun);
END_METHOD

{region 'Documentation'}
(*!
<summary>Returns a registered scenario using its original array index.</summary>
*)
{endregion}
METHOD PUBLIC GetTestCase : I_TestCase //! Typed child interface at the original array index; zero when no entry is available.
VAR_INPUT
    Index : DINT; //! Original occupied child-array index, rather than an ordinal position.
END_VAR
GetTestCase := 0;
IF (ChildCount = 0) OR (Index < ChildArrayLowerBound)
    OR (DINT_TO_LINT(Index) >= DINT_TO_LINT(ChildArrayLowerBound) + UINT_TO_LINT(ChildCount)) THEN
    RETURN;
END_IF;
GetTestCase := FTestCases[Index];
END_METHOD

{region 'Documentation'}
(*!
<summary>Calls each owned scenario once per initialized Suite cycle.</summary>
*)
{endregion}
METHOD PROTECTED ProcessTestCases
FEpochs();
FCommands();
FActiveRun();
END_METHOD

END_FUNCTION_BLOCK

// ---- SelfTests/TestCases/TestSuite_EventBufferReset/Test_BufferResetEpochs.TcPOU
{region 'Documentation'}
(*!
<summary>Checks coordinated hard reset of empty, populated and full wrapped local Event Buffer epochs.</summary>
<description>
RunControlIntegrationSubject executes the real hierarchy once per test cycle until Idle.
Each scenario reserves through the actual Suite and Test Cases before arranging its buffer.
Only ControlData.BufferCmd.Reset requests a hard reset; setup uses ordinary publication and deletion.
The Idle subject must not publish a reset-only event or change lifecycle. Checks accumulate across
all three scenarios, including typed empty fields in every physical ring position and sequence restart.
The full wrapped scenario deliberately fills reserved capacity and loses one event as reset input;
this tests destructive recovery, not normal admission or a promise of loss-free publication.
The real subject binds only local storage; expected findings remain in that storage.
Checking Assertions retain the outer selftest publisher. Each run reinitializes the subject.
</description>
*)
{endregion}
FUNCTION_BLOCK Test_BufferResetEpochs EXTENDS TestCaseBase
VAR
    FSubject : EventBuffer;
    FEvents : ARRAY[1..BufferLength] OF ST_Event;
    FFifo : ST_FifoStatus;
    FBufferStatus : ST_EventBufferStatus;
    FPerformed : BOOL;
    FChecked : BOOL;
    FRoot : RunControlIntegrationSubject;
    FControl : ST_RunControl;
    FPhase : USINT;
    FScenario : USINT;
    FScenarioPrepared : BOOL;
    FSuite : I_TestSuite;
    FFirstChild : I_TestCase;
    FSecondChild : I_TestCase;
    FSetup : AssertTrue;
    FSetupMatches : BOOL;
    FEmptyEpoch : AssertTrue;
    FEmptyEpochMatches : BOOL;
    FFilledEpoch : AssertTrue;
    FFilledEpochMatches : BOOL;
    FWrappedEpoch : AssertTrue;
    FWrappedEpochMatches : BOOL;
    FStorageCleared : AssertTrue;
    FStorageClearedMatches : BOOL;
    FReservationsReleased : AssertTrue;
    FReservationsReleasedMatches : BOOL;
    FCommandClearing : AssertTrue;
    FCommandClearingMatches : BOOL;
    FLifecyclePreserved : AssertTrue;
    FLifecyclePreservedMatches : BOOL;
    FNewEpoch : AssertTrue;
    FNewEpochMatches : BOOL;
END_VAR
VAR CONSTANT
    BufferLength : UINT := 129;
    SeedEventCount : UINT := 6;
    DeletedSeedCount : UDINT := 4;
    EmptyScenario : USINT := 0;
    FilledScenario : USINT := 1;
    WrappedScenario : USINT := 2;
    SetupPhase : USINT := 0;
    AwaitIdlePhase : USINT := 1;
    PreparePhase : USINT := 2;
    ResetPhase : USINT := 3;
    VerifyPhase : USINT := 4;
END_VAR

SUPER^();

{region 'Documentation'}
(*!
<summary>Contributes each checking Assertion once.</summary>
*)
{endregion}
METHOD PROTECTED AggregateResults
VAR_INPUT
    Aggregator : I_ResultAggregator; //! Borrowed result sink owned by the outer Test Case; add this test's checking Assertions without resetting or retaining the sink.
END_VAR
Aggregator.AddProvider(Provider := FSetup);
Aggregator.AddProvider(Provider := FEmptyEpoch);
Aggregator.AddProvider(Provider := FFilledEpoch);
Aggregator.AddProvider(Provider := FWrappedEpoch);
Aggregator.AddProvider(Provider := FStorageCleared);
Aggregator.AddProvider(Provider := FReservationsReleased);
Aggregator.AddProvider(Provider := FCommandClearing);
Aggregator.AddProvider(Provider := FLifecyclePreserved);
Aggregator.AddProvider(Provider := FNewEpoch);
END_METHOD

{region 'Documentation'}
(*!
<summary>Requires all checking Assertions to be initialized.</summary>
*)
{endregion}
METHOD PROTECTED CheckInitialization : BOOL //! TRUE when the inherited initialization check and this concrete fixture check both accept the setup.
CheckInitialization := FALSE;
IF NOT SUPER^.CheckInitialization() THEN
    RETURN;
END_IF;

CheckInitialization := FSetup.IsInitialized
    AND FEmptyEpoch.IsInitialized
    AND FFilledEpoch.IsInitialized
    AND FWrappedEpoch.IsInitialized
    AND FStorageCleared.IsInitialized
    AND FReservationsReleased.IsInitialized
    AND FCommandClearing.IsInitialized
    AND FLifecyclePreserved.IsInitialized
    AND FNewEpoch.IsInitialized;
END_METHOD

{region 'Documentation'}
(*!
<summary>Checks typed empty storage, epoch metadata and real hierarchical release after the root call.</summary>
*)
{endregion}
METHOD PRIVATE CheckReset
VAR
    Index : UINT;
    EmptyEvent : ST_Event;
    EpochCleared : BOOL;
END_VAR
EpochCleared := FFifo.BufferEmpty AND NOT FFifo.BufferFull AND NOT FFifo.BufferAlmostFull
    AND (FFifo.ElementCount = 0) AND (FFifo.BufferLength = BufferLength)
    AND (FFifo.IndexIn = 1) AND (FFifo.IndexOut = 1)
    AND NOT FFifo.ConfigError AND NOT FFifo.IndexError
    AND (FBufferStatus.SequenceId = 0) AND (FBufferStatus.DeletedSequenceId = 0)
    AND (FBufferStatus.LostEventCount = 0);
CASE FScenario OF
    EmptyScenario:
        FEmptyEpochMatches := FScenarioPrepared AND EpochCleared;
    FilledScenario:
        FFilledEpochMatches := FScenarioPrepared AND EpochCleared;
    WrappedScenario:
        FWrappedEpochMatches := FScenarioPrepared AND EpochCleared;
    ELSE
        Error(Message := 'Unknown local reset observation scenario.');
END_CASE;

FOR Index := 1 TO BufferLength DO
    FStorageClearedMatches := FStorageClearedMatches
        AND (FEvents[Index].SequenceId = EmptyEvent.SequenceId)
        AND (FEvents[Index].Timestamp = EmptyEvent.Timestamp)
        AND (FEvents[Index].OwnerScope = EmptyEvent.OwnerScope)
        AND (FEvents[Index].EventType = EmptyEvent.EventType)
        AND (FEvents[Index].Severity = EmptyEvent.Severity)
        AND (FEvents[Index].Name = EmptyEvent.Name)
        AND (FEvents[Index].ResourceName = EmptyEvent.ResourceName)
        AND (FEvents[Index].State = EmptyEvent.State)
        AND (FEvents[Index].Result = EmptyEvent.Result)
        AND (FEvents[Index].Message = EmptyEvent.Message);
END_FOR;
FReservationsReleasedMatches := FReservationsReleasedMatches
    AND (FSubject.ReservedEntryCount = 0) AND (FSuite.ReservedEntryCount = 0)
    AND (FFirstChild.ReservedEntryCount = 0) AND (FSecondChild.ReservedEntryCount = 0);
FCommandClearingMatches := FCommandClearingMatches
    AND NOT FControl.BufferCmd.Reset AND (FControl.BufferCmd.DeleteSequenceId = 0);
FLifecyclePreservedMatches := FLifecyclePreservedMatches AND FRoot.IsIdle AND FRoot.IsReady
    AND (FSuite.State = E_State.Idle) AND (FFirstChild.State = E_State.Idle)
    AND (FSecondChild.State = E_State.Idle) AND FRoot.ConfigurationUnchanged
    AND FRoot.ChildCallsMatch;
END_METHOD

{region 'Documentation'}
(*!
<summary>Initializes the checking Assertions for one test state.</summary>
*)
{endregion}
METHOD PROTECTED Configure
FPreparationStateCount := 0;
FTestStateCount := 1;
FSetup.Initialize(Parent := THIS^,
    AssertionName := 'Setup');
FEmptyEpoch.Initialize(Parent := THIS^,
    AssertionName := 'EmptyEpoch');
FFilledEpoch.Initialize(Parent := THIS^,
    AssertionName := 'FilledEpoch');
FWrappedEpoch.Initialize(Parent := THIS^,
    AssertionName := 'WrappedEpoch');
FStorageCleared.Initialize(Parent := THIS^,
    AssertionName := 'StorageCleared');
FReservationsReleased.Initialize(Parent := THIS^,
    AssertionName := 'ReservationsReleased');
FCommandClearing.Initialize(Parent := THIS^,
    AssertionName := 'CommandClearing');
FLifecyclePreserved.Initialize(Parent := THIS^,
    AssertionName := 'LifecyclePreserved');
FNewEpoch.Initialize(Parent := THIS^,
    AssertionName := 'NewEpoch');
END_METHOD

{region 'Documentation'}
(*!
<summary>Builds a known epoch through real Publish/Delete calls and owner reservation methods.</summary>
*)
{endregion}
METHOD PRIVATE PrepareScenario
VAR
    Index : UINT;
    SequenceBefore : UDINT;
    Published : INT;
    SuiteReservation : E_EventReservationResult;
    FirstReservation : E_EventReservationResult;
    SecondReservation : E_EventReservationResult;
    SeedEvent : ST_Event;
END_VAR
FControl.BufferCmd.DeleteSequenceId := FBufferStatus.SequenceId;
FSubject.ProcessDeleteRequest(SequenceId := FControl.BufferCmd.DeleteSequenceId);
SuiteReservation := FSuite.ReserveResetEvents();
FirstReservation := FFirstChild.ReserveResetEvents();
SecondReservation := FSecondChild.ReserveResetEvents();
FSetupMatches := FSetupMatches AND FFifo.BufferEmpty
    AND (SuiteReservation = E_EventReservationResult.Accepted)
    AND (FirstReservation = E_EventReservationResult.Accepted)
    AND (SecondReservation = E_EventReservationResult.Accepted)
    AND (FSuite.ReservedEntryCount = GVL_Constants.TestSuiteResetEventCount)
    AND (FFirstChild.ReservedEntryCount = GVL_Constants.TestCaseResetEventCount)
    AND (FSecondChild.ReservedEntryCount = GVL_Constants.TestCaseResetEventCount)
    AND (FSubject.ReservedEntryCount = GVL_Constants.TestSuiteResetEventCount
        + 2 * GVL_Constants.TestCaseResetEventCount);
SeedEvent := CreateFrameworkEvent(Name := 'ResetSubject',
    ResourceName := 'ResetFixture',
    State := E_State.Idle,
    Severity := E_EventSeverity.Info,
    Message := 'Discarded by coordinated hard reset.');
SequenceBefore := FBufferStatus.SequenceId;

CASE FScenario OF
    EmptyScenario:
        FScenarioPrepared := FFifo.BufferEmpty
            AND (FBufferStatus.SequenceId = FBufferStatus.DeletedSequenceId)
            AND (FBufferStatus.LostEventCount = 0);

    FilledScenario, WrappedScenario:
        FOR Index := 1 TO SeedEventCount DO
            Published := FSubject.PublishEvent(Event := SeedEvent);
            FSetupMatches := FSetupMatches AND (Published > 0);
        END_FOR;
        FControl.BufferCmd.DeleteSequenceId := SequenceBefore + DeletedSeedCount;
        FSubject.ProcessDeleteRequest(SequenceId := FControl.BufferCmd.DeleteSequenceId);
        FScenarioPrepared := (FFifo.ElementCount = SeedEventCount - UDINT_TO_UINT(DeletedSeedCount))
            AND (FBufferStatus.SequenceId = SequenceBefore + UINT_TO_UDINT(SeedEventCount))
            AND (FBufferStatus.DeletedSequenceId = SequenceBefore + DeletedSeedCount)
            AND (FBufferStatus.LostEventCount = 0);
        IF FScenario = WrappedScenario THEN
            FOR Index := 1 TO BufferLength DO
                IF FFifo.BufferFull THEN
                    EXIT;
                END_IF;
                Published := FSubject.PublishEvent(Event := SeedEvent);
                FSetupMatches := FSetupMatches AND (Published > 0);
            END_FOR;
            SequenceBefore := FBufferStatus.SequenceId;
            Published := FSubject.PublishEvent(Event := SeedEvent);
            FScenarioPrepared := FScenarioPrepared AND FFifo.BufferFull
                AND (FFifo.ElementCount = BufferLength - 1) AND (FFifo.IndexIn < FFifo.IndexOut)
                AND (Published = TO_INT(E_FifoResult.NoTransfer))
                AND (FBufferStatus.SequenceId = SequenceBefore + 1)
                AND (FBufferStatus.LostEventCount = 1);
        END_IF;

    ELSE
        Error(Message := 'Unknown local buffer epoch scenario.');
END_CASE;
END_METHOD

{region 'Documentation'}
(*!
<summary>Completes abort without asynchronous work.</summary>
*)
{endregion}
METHOD PROTECTED ProcessAbort
VAR_INPUT
    Enable : BOOL; //! Phase permission supplied by the owning Test Case; FALSE does not authorize progression, while observation may continue.
END_VAR
IF Enable THEN
    CompleteAbort();
END_IF;
END_METHOD

{region 'Documentation'}
(*!
<summary>Evaluates captured observations after the scenario has finished.</summary>
*)
{endregion}
METHOD PROTECTED ProcessAssertions
VAR_INPUT
    Enable : BOOL; //! Phase permission supplied by the owning Test Case; FALSE does not authorize progression, while observation may continue.
END_VAR
VAR
    Evaluate : BOOL;
END_VAR
Evaluate := Enable AND FPerformed;
FSetup(Enable := Evaluate,
    State := State,
    IN := FSetupMatches);
FEmptyEpoch(Enable := Evaluate,
    State := State,
    IN := FEmptyEpochMatches);
FFilledEpoch(Enable := Evaluate,
    State := State,
    IN := FFilledEpochMatches);
FWrappedEpoch(Enable := Evaluate,
    State := State,
    IN := FWrappedEpochMatches);
FStorageCleared(Enable := Evaluate,
    State := State,
    IN := FStorageClearedMatches);
FReservationsReleased(Enable := Evaluate,
    State := State,
    IN := FReservationsReleasedMatches);
FCommandClearing(Enable := Evaluate,
    State := State,
    IN := FCommandClearingMatches);
FLifecyclePreserved(Enable := Evaluate,
    State := State,
    IN := FLifecyclePreservedMatches);
FNewEpoch(Enable := Evaluate,
    State := State,
    IN := FNewEpochMatches);
IF Evaluate THEN
    FChecked := TRUE;
END_IF;
END_METHOD

{region 'Documentation'}
(*!
<summary>No Preparation phase is needed.</summary>
*)
{endregion}
METHOD PROTECTED ProcessPreparations
VAR_INPUT
    // SA0033: Required override without Preparation work.
    {attribute 'analysis' := '-33'}
    Enable : BOOL; //! Phase permission supplied by the owning Test Case; FALSE does not authorize progression, while observation may continue.
END_VAR
END_METHOD

{region 'Documentation'}
(*!
<summary>Resets observations and schedules a fresh subject initialization.</summary>
*)
{endregion}
METHOD PROTECTED ProcessReset
FPerformed := FALSE;
FChecked := FALSE;
FPhase := SetupPhase;
FScenario := EmptyScenario;
FScenarioPrepared := FALSE;
FSuite := 0;
FFirstChild := 0;
FSecondChild := 0;
FSetup.Reset();
FSetupMatches := TRUE;
FEmptyEpoch.Reset();
FEmptyEpochMatches := TRUE;
FFilledEpoch.Reset();
FFilledEpochMatches := TRUE;
FWrappedEpoch.Reset();
FWrappedEpochMatches := TRUE;
FStorageCleared.Reset();
FStorageClearedMatches := TRUE;
FReservationsReleased.Reset();
FReservationsReleasedMatches := TRUE;
FCommandClearing.Reset();
FCommandClearingMatches := TRUE;
FLifecyclePreserved.Reset();
FLifecyclePreservedMatches := TRUE;
FNewEpoch.Reset();
FNewEpochMatches := TRUE;
CompleteReset();
END_METHOD

{region 'Documentation'}
(*!
<summary>Advances one scenario phase per PLC cycle before evaluating accumulated checks.</summary>
*)
{endregion}
METHOD PROTECTED ProcessTests
VAR_INPUT
    Enable : BOOL; //! Phase permission supplied by the owning Test Case; FALSE does not authorize progression, while observation may continue.
END_VAR
IF NOT Enable THEN
    RETURN;
END_IF;
IF FChecked THEN
    CompleteTests();
    RETURN;
END_IF;

IF NOT FPerformed THEN
    StateMachine();
END_IF;
END_METHOD

{region 'Documentation'}
(*!
<summary>Executes one subject call per active test cycle; all reset observations follow that call.</summary>
*)
{endregion}
METHOD PRIVATE StateMachine
VAR
    EmptyControl : ST_RunControl;
END_VAR
CASE FPhase OF
    SetupPhase:
        FControl := EmptyControl;
        IF NOT FSubject.Initialize(Buffer := FEvents,
            FifoControl := FFifo,
            Status := FBufferStatus) THEN
            Error(Message := 'Local reset buffer initialization failed.');
            RETURN;
        END_IF;
        FRoot.BindPublisher(Publisher := FSubject);
        IF NOT FRoot.Initialize(Name := 'ResetSubject',
            EventBuffer := FSubject) THEN
            Error(Message := 'Local reset root initialization failed.');
            RETURN;
        END_IF;
        FPhase := AwaitIdlePhase;

    AwaitIdlePhase:
        FRoot(ControlData := FControl);
        IF FRoot.HasError THEN
            Error(Message := 'Local hierarchy did not establish the Idle reset precondition.');
            RETURN;
        END_IF;
        IF FRoot.IsReady THEN
            FSuite := FRoot.GetTestSuite(Index := FRoot.ChildArrayLowerBound);
            FFirstChild := FRoot.GetTestCase(Index := FRoot.TestCaseLowerBound);
            FSecondChild := FRoot.GetTestCase(Index := FRoot.TestCaseLowerBound + 1);
            IF (FSuite = 0) OR (FFirstChild = 0) OR (FSecondChild = 0) THEN
                Error(Message := 'Local reset hierarchy has missing registered children.');
                RETURN;
            END_IF;
            FPhase := PreparePhase;
        END_IF;

    PreparePhase:
        FRoot(ControlData := FControl);
        PrepareScenario();
        FPhase := ResetPhase;

    ResetPhase:
        FControl.BufferCmd.Reset := TRUE;
        FRoot(ControlData := FControl);
        CheckReset();
        FPhase := VerifyPhase;

    VerifyPhase:
        VerifyNewEpoch();
        FRoot(ControlData := FControl);
        FLifecyclePreservedMatches := FLifecyclePreservedMatches AND FRoot.IsIdle
            AND FRoot.IsReady AND FRoot.ConfigurationUnchanged AND FRoot.ChildCallsMatch;
        IF FScenario = WrappedScenario THEN
            FPerformed := TRUE;
        ELSE
            FScenario := FScenario + 1;
            FPhase := PreparePhase;
        END_IF;

    ELSE
        Error(Message := 'Unknown local buffer reset scenario phase.');
END_CASE;
END_METHOD

{region 'Documentation'}
(*!
<summary>Publishes the first new event and checks sequence restart without old payload retention.</summary>
*)
{endregion}
METHOD PRIVATE VerifyNewEpoch
VAR
    Published : INT;
END_VAR
Published := FSubject.PublishEvent(Event := CreateFrameworkEvent(Name := 'ResetSubject',
    State := E_State.Idle,
    Severity := E_EventSeverity.Info,
    Message := 'First event in the new epoch.'));
FNewEpochMatches := FNewEpochMatches AND (Published > 0)
    AND (FBufferStatus.SequenceId = 1) AND (FBufferStatus.DeletedSequenceId = 0)
    AND (FBufferStatus.LostEventCount = 0) AND (FFifo.ElementCount = 1)
    AND (FEvents[FFifo.IndexOut].SequenceId = 1)
    AND (FEvents[FFifo.IndexOut].Message = 'First event in the new epoch.');
END_METHOD

END_FUNCTION_BLOCK

// ---- SelfTests/TestCases/TestSuite_EventBufferReset/Test_BufferResetCommands.TcPOU
{region 'Documentation'}
(*!
<summary>Checks reset/delete priority, release ordering and destructive reset after a controlled Suite release failure.</summary>
<description>
Two scenarios use successful releases, then a rejected first Suite release followed by a successful second.
A real Event Buffer probe records release/reset ordering and nonzero delete submissions.
The controlled Orchestrator keeps lifecycle Idle and cannot conceal command work with its own releases.
The failed Suite contribution intentionally remains; only the hard-reset buffer aggregate is guaranteed clear.
The real subject binds only local storage; expected findings remain in that storage.
Checking Assertions retain the outer selftest publisher. Each run reinitializes the subject.
</description>
*)
{endregion}
FUNCTION_BLOCK Test_BufferResetCommands EXTENDS TestCaseBase
VAR
    FSubject : BufferCommandProbe;
    FEvents : ARRAY[1..BufferLength] OF ST_Event;
    FFifo : ST_FifoStatus;
    FBufferStatus : ST_EventBufferStatus;
    FPerformed : BOOL;
    FChecked : BOOL;
    FRoot : BufferResetRunControlProbe;
    FHelper : SuiteOrchestratorDouble;
    FFirstSuite : BufferReleaseSuiteDouble;
    FSecondSuite : BufferReleaseSuiteDouble;
    FControl : ST_RunControl;
    FPhase : USINT;
    FRejectFirstRelease : BOOL;
    FSetup : AssertTrue;
    FSetupMatches : BOOL;
    FDeleteOnly : AssertTrue;
    FDeleteOnlyMatches : BOOL;
    FResetPriority : AssertTrue;
    FResetPriorityMatches : BOOL;
    FReleaseOrder : AssertTrue;
    FReleaseOrderMatches : BOOL;
    FReleaseFailure : AssertTrue;
    FReleaseFailureMatches : BOOL;
    FHardReset : AssertTrue;
    FHardResetMatches : BOOL;
    FCommandsCleared : AssertTrue;
    FCommandsClearedMatches : BOOL;
    FNoReplay : AssertTrue;
    FNoReplayMatches : BOOL;
    FLifecyclePreserved : AssertTrue;
    FLifecyclePreservedMatches : BOOL;
END_VAR
VAR CONSTANT
    BufferLength : UINT := 65;
    Contribution : UINT := 3;
    SetupPhase : USINT := 0;
    AwaitIdlePhase : USINT := 1;
    DeletePhase : USINT := 2;
    PreparePhase : USINT := 3;
    ResetPhase : USINT := 4;
    VerifyPhase : USINT := 5;
END_VAR

SUPER^();

{region 'Documentation'}
(*!
<summary>Contributes each checking Assertion once.</summary>
*)
{endregion}
METHOD PROTECTED AggregateResults
VAR_INPUT
    Aggregator : I_ResultAggregator; //! Borrowed result sink owned by the outer Test Case; add this test's checking Assertions without resetting or retaining the sink.
END_VAR
Aggregator.AddProvider(Provider := FSetup);
Aggregator.AddProvider(Provider := FDeleteOnly);
Aggregator.AddProvider(Provider := FResetPriority);
Aggregator.AddProvider(Provider := FReleaseOrder);
Aggregator.AddProvider(Provider := FReleaseFailure);
Aggregator.AddProvider(Provider := FHardReset);
Aggregator.AddProvider(Provider := FCommandsCleared);
Aggregator.AddProvider(Provider := FNoReplay);
Aggregator.AddProvider(Provider := FLifecyclePreserved);
END_METHOD

{region 'Documentation'}
(*!
<summary>Requires all checking Assertions to be initialized.</summary>
*)
{endregion}
METHOD PROTECTED CheckInitialization : BOOL //! TRUE when the inherited initialization check and this concrete fixture check both accept the setup.
CheckInitialization := FALSE;
IF NOT SUPER^.CheckInitialization() THEN
    RETURN;
END_IF;

CheckInitialization := FSetup.IsInitialized
    AND FDeleteOnly.IsInitialized
    AND FResetPriority.IsInitialized
    AND FReleaseOrder.IsInitialized
    AND FReleaseFailure.IsInitialized
    AND FHardReset.IsInitialized
    AND FCommandsCleared.IsInitialized
    AND FNoReplay.IsInitialized
    AND FLifecyclePreserved.IsInitialized;
END_METHOD

{region 'Documentation'}
(*!
<summary>Initializes the checking Assertions for one test state.</summary>
*)
{endregion}
METHOD PROTECTED Configure
FPreparationStateCount := 0;
FTestStateCount := 1;
FSetup.Initialize(Parent := THIS^,
    AssertionName := 'Setup');
FDeleteOnly.Initialize(Parent := THIS^,
    AssertionName := 'DeleteOnly');
FResetPriority.Initialize(Parent := THIS^,
    AssertionName := 'ResetPriority');
FReleaseOrder.Initialize(Parent := THIS^,
    AssertionName := 'ReleaseOrder');
FReleaseFailure.Initialize(Parent := THIS^,
    AssertionName := 'ReleaseFailure');
FHardReset.Initialize(Parent := THIS^,
    AssertionName := 'HardReset');
FCommandsCleared.Initialize(Parent := THIS^,
    AssertionName := 'CommandsCleared');
FNoReplay.Initialize(Parent := THIS^,
    AssertionName := 'NoReplay');
FLifecyclePreserved.Initialize(Parent := THIS^,
    AssertionName := 'LifecyclePreserved');
END_METHOD

{region 'Documentation'}
(*!
<summary>Creates a populated epoch and real contributions before starting order observation.</summary>
*)
{endregion}
METHOD PRIVATE PrepareReset
VAR
    SeedEvent : ST_Event;
    Published : INT;
    FirstReserved : BOOL;
    SecondReserved : BOOL;
END_VAR
SeedEvent := CreateFrameworkEvent(Name := 'ResetCommands',
    ResourceName := 'CommandFixture',
    State := E_State.Idle,
    Severity := E_EventSeverity.Info,
    Message := 'Pending deletion must be superseded by hard reset.');
Published := FSubject.PublishEvent(Event := SeedEvent);
FirstReserved := FFirstSuite.PrepareRelease(RejectRelease := FRejectFirstRelease,
    EntryCount := Contribution,
    Buffer := FSubject);
SecondReserved := FSecondSuite.PrepareRelease(RejectRelease := FALSE,
    EntryCount := Contribution,
    Buffer := FSubject);
FSetupMatches := FSetupMatches AND (Published > 0) AND FirstReserved AND SecondReserved
    AND (FSubject.ReservedEntryCount = 2 * Contribution) AND NOT FFifo.BufferEmpty;
FFirstSuite.BeginCycle();
FSecondSuite.BeginCycle();
FSubject.BeginObservation();
END_METHOD

{region 'Documentation'}
(*!
<summary>Completes abort without asynchronous work.</summary>
*)
{endregion}
METHOD PROTECTED ProcessAbort
VAR_INPUT
    Enable : BOOL; //! Phase permission supplied by the owning Test Case; FALSE does not authorize progression, while observation may continue.
END_VAR
IF Enable THEN
    CompleteAbort();
END_IF;
END_METHOD

{region 'Documentation'}
(*!
<summary>Evaluates captured observations after the scenario has finished.</summary>
*)
{endregion}
METHOD PROTECTED ProcessAssertions
VAR_INPUT
    Enable : BOOL; //! Phase permission supplied by the owning Test Case; FALSE does not authorize progression, while observation may continue.
END_VAR
VAR
    Evaluate : BOOL;
END_VAR
Evaluate := Enable AND FPerformed;
FSetup(Enable := Evaluate,
    State := State,
    IN := FSetupMatches);
FDeleteOnly(Enable := Evaluate,
    State := State,
    IN := FDeleteOnlyMatches);
FResetPriority(Enable := Evaluate,
    State := State,
    IN := FResetPriorityMatches);
FReleaseOrder(Enable := Evaluate,
    State := State,
    IN := FReleaseOrderMatches);
FReleaseFailure(Enable := Evaluate,
    State := State,
    IN := FReleaseFailureMatches);
FHardReset(Enable := Evaluate,
    State := State,
    IN := FHardResetMatches);
FCommandsCleared(Enable := Evaluate,
    State := State,
    IN := FCommandsClearedMatches);
FNoReplay(Enable := Evaluate,
    State := State,
    IN := FNoReplayMatches);
FLifecyclePreserved(Enable := Evaluate,
    State := State,
    IN := FLifecyclePreservedMatches);
IF Evaluate THEN
    FChecked := TRUE;
END_IF;
END_METHOD

{region 'Documentation'}
(*!
<summary>No Preparation phase is needed.</summary>
*)
{endregion}
METHOD PROTECTED ProcessPreparations
VAR_INPUT
    // SA0033: Required override without Preparation work.
    {attribute 'analysis' := '-33'}
    Enable : BOOL; //! Phase permission supplied by the owning Test Case; FALSE does not authorize progression, while observation may continue.
END_VAR
END_METHOD

{region 'Documentation'}
(*!
<summary>Resets observations and schedules a fresh subject initialization.</summary>
*)
{endregion}
METHOD PROTECTED ProcessReset
FPerformed := FALSE;
FChecked := FALSE;
FPhase := SetupPhase;
FRejectFirstRelease := FALSE;
FSetup.Reset();
FSetupMatches := TRUE;
FDeleteOnly.Reset();
FDeleteOnlyMatches := TRUE;
FResetPriority.Reset();
FResetPriorityMatches := TRUE;
FReleaseOrder.Reset();
FReleaseOrderMatches := TRUE;
FReleaseFailure.Reset();
FReleaseFailureMatches := TRUE;
FHardReset.Reset();
FHardResetMatches := TRUE;
FCommandsCleared.Reset();
FCommandsClearedMatches := TRUE;
FNoReplay.Reset();
FNoReplayMatches := TRUE;
FLifecyclePreserved.Reset();
FLifecyclePreservedMatches := TRUE;
CompleteReset();
END_METHOD

{region 'Documentation'}
(*!
<summary>Runs the bounded scenario once before Assertion evaluation.</summary>
*)
{endregion}
METHOD PROTECTED ProcessTests
VAR_INPUT
    Enable : BOOL; //! Phase permission supplied by the owning Test Case; FALSE does not authorize progression, while observation may continue.
END_VAR
IF NOT Enable THEN
    RETURN;
END_IF;
IF FChecked THEN
    CompleteTests();
    RETURN;
END_IF;

IF NOT FPerformed THEN
    StateMachine();
END_IF;
END_METHOD

{region 'Documentation'}
(*!
<summary>Advances one owner call per cycle and records command observations immediately after it.</summary>
*)
{endregion}
METHOD PRIVATE StateMachine
VAR
    EmptyControl : ST_RunControl;
    SeedEvent : ST_Event;
    Published : INT;
    FirstCalls : ST_OrchestrationCalls;
    SecondCalls : ST_OrchestrationCalls;
END_VAR
CASE FPhase OF
    SetupPhase:
        FControl := EmptyControl;
        IF NOT FSubject.Initialize(Buffer := FEvents,
            FifoControl := FFifo,
            Status := FBufferStatus) THEN
            Error(Message := 'Command-test buffer initialization failed.');
            RETURN;
        END_IF;
        FHelper.BeginScenario();
        FRoot.Bind(Publisher := FSubject,
            Helper := FHelper);
        FRoot.BindChildren(FirstSuite := FFirstSuite,
            SecondSuite := FSecondSuite);
        IF NOT FRoot.Initialize(Name := 'ResetCommands',
            EventBuffer := FSubject) THEN
            Error(Message := 'Command-test root initialization failed.');
            RETURN;
        END_IF;
        FHelper.SetObservation(Ready := TRUE,
            ResetFinished := TRUE);
        FPhase := AwaitIdlePhase;

    AwaitIdlePhase:
        FRoot(ControlData := FControl);
        IF FRoot.HasError THEN
            Error(Message := 'Command-test root did not establish Idle.');
            RETURN;
        END_IF;
        IF FRoot.IsReady THEN
            FSubject.BeginObservation();
            FControl.BufferCmd.DeleteSequenceId := FBufferStatus.SequenceId;
            FSetupMatches := FSetupMatches AND (FControl.BufferCmd.DeleteSequenceId > 0);
            FPhase := DeletePhase;
        END_IF;

    DeletePhase:
        FRoot(ControlData := FControl);
        FDeleteOnlyMatches := (FSubject.DeleteCount = 1) AND (FSubject.ResetCount = 0)
            AND FFifo.BufferEmpty AND (FControl.BufferCmd.DeleteSequenceId = 0)
            AND (FBufferStatus.DeletedSequenceId = FBufferStatus.SequenceId);
        FPhase := PreparePhase;

    PreparePhase:
        FRoot(ControlData := FControl);
        PrepareReset();
        FPhase := ResetPhase;

    ResetPhase:
        FControl.BufferCmd.Reset := TRUE;
        FControl.BufferCmd.DeleteSequenceId := FBufferStatus.SequenceId;
        FRoot(ControlData := FControl);
        FResetPriorityMatches := FResetPriorityMatches AND (FSubject.DeleteCount = 0)
            AND (FSubject.ResetCount = 1);
        FReleaseOrderMatches := FReleaseOrderMatches
            AND (FFirstSuite.ReleaseCount = 1) AND (FSecondSuite.ReleaseCount = 1)
            AND (FFirstSuite.ReleaseOrder = 1) AND (FSecondSuite.ReleaseOrder = 2)
            AND (FSubject.ResetOrder = 3);
        FReleaseFailureMatches := FReleaseFailureMatches AND (FSecondSuite.ReservedEntryCount = 0);
        IF FRejectFirstRelease THEN
            FReleaseFailureMatches := FReleaseFailureMatches
                AND (FFirstSuite.ReservedEntryCount = Contribution);
        ELSE
            FReleaseFailureMatches := FReleaseFailureMatches
                AND (FFirstSuite.ReservedEntryCount = 0);
        END_IF;
        FHardResetMatches := FHardResetMatches AND FFifo.BufferEmpty
            AND (FFifo.ElementCount = 0) AND (FBufferStatus.SequenceId = 0)
            AND (FBufferStatus.DeletedSequenceId = 0) AND (FBufferStatus.LostEventCount = 0)
            AND (FSubject.ReservedEntryCount = 0);
        FCommandsClearedMatches := FCommandsClearedMatches AND NOT FControl.BufferCmd.Reset
            AND (FControl.BufferCmd.DeleteSequenceId = 0);
        FirstCalls := FFirstSuite.Calls;
        SecondCalls := FSecondSuite.Calls;
        FLifecyclePreservedMatches := FLifecyclePreservedMatches AND FRoot.IsIdle AND FRoot.IsReady
            AND (FFirstSuite.State = E_State.Idle) AND (FSecondSuite.State = E_State.Idle)
            AND (FirstCalls.ResetCount = 0) AND (FirstCalls.StartCount = 0)
            AND (FirstCalls.AbortCount = 0) AND (SecondCalls.ResetCount = 0)
            AND (SecondCalls.StartCount = 0) AND (SecondCalls.AbortCount = 0);
        FPhase := VerifyPhase;

    VerifyPhase:
        SeedEvent := CreateFrameworkEvent(Name := 'ResetCommands',
            ResourceName := 'CommandFixture',
            State := E_State.Idle,
            Severity := E_EventSeverity.Info,
            Message := 'New epoch must survive the next owner call.');
        Published := FSubject.PublishEvent(Event := SeedEvent);
        FRoot(ControlData := FControl);
        FNoReplayMatches := FNoReplayMatches AND (Published > 0)
            AND (FSubject.ResetCount = 1) AND (FSubject.DeleteCount = 0)
            AND (FFirstSuite.ReleaseCount = 1) AND (FSecondSuite.ReleaseCount = 1)
            AND (FBufferStatus.SequenceId = 1) AND (FFifo.ElementCount = 1);
        IF FRejectFirstRelease THEN
            FPerformed := TRUE;
        ELSE
            FRejectFirstRelease := TRUE;
            FPhase := PreparePhase;
        END_IF;

    ELSE
        Error(Message := 'Unknown buffer command-test phase.');
END_CASE;
END_METHOD

END_FUNCTION_BLOCK

// ---- SelfTests/TestCases/TestSuite_EventBufferReset/Helper/BufferCommandProbe.TcPOU
{region 'Documentation'}
(*!
<summary>Real Event Buffer with command-order observations; BeginObservation excludes setup calls.</summary>
*)
{endregion}
FUNCTION_BLOCK BufferCommandProbe EXTENDS EventBuffer
VAR
    FOperationCount : UINT;
    FResetOrder : UINT;
    FResetCount : UINT;
    FDeleteCount : UINT;
END_VAR

{region 'Documentation'}
(*!
<summary>Clears only test observations, not buffer contents or reservations.</summary>
*)
{endregion}
METHOD PUBLIC BeginObservation
FOperationCount := 0;
FResetOrder := 0;
FResetCount := 0;
FDeleteCount := 0;
END_METHOD

{region 'Documentation'}
(*!
<summary>Recorded DeleteCount for command-order verification.</summary>
*)
{endregion}
{attribute 'monitoring' := 'call'}
PROPERTY PUBLIC DeleteCount : UINT //! Recorded DeleteCount for command-order verification.
GET
DeleteCount := FDeleteCount;
END_GET
END_PROPERTY

{region 'Documentation'}
(*!
<summary>Counts nonzero delete commands, then delegates unchanged to the real buffer.</summary>
*)
{endregion}
METHOD PUBLIC ProcessDeleteRequest
VAR_IN_OUT
    SequenceId : UDINT; //! Pending delete watermark passed through to the inherited consumer, which clears the request.
END_VAR
IF SequenceId <> 0 THEN
    FDeleteCount := FDeleteCount + 1;
END_IF;
SUPER^.ProcessDeleteRequest(SequenceId := SequenceId);
END_METHOD

{region 'Documentation'}
(*!
<summary>Records a Suite release attempt in the same order domain as Reset.</summary>
*)
{endregion}
METHOD PUBLIC RecordRelease : UINT //! Incremented operation sequence number shared with buffer Reset observations.
FOperationCount := FOperationCount + 1;
RecordRelease := FOperationCount;
END_METHOD

{region 'Documentation'}
(*!
<summary>Records entry, then executes the unchanged real hard reset.</summary>
*)
{endregion}
METHOD PUBLIC Reset
FOperationCount := FOperationCount + 1;
FResetOrder := FOperationCount;
FResetCount := FResetCount + 1;
SUPER^.Reset();
END_METHOD

{region 'Documentation'}
(*!
<summary>Recorded ResetCount for command-order verification.</summary>
*)
{endregion}
{attribute 'monitoring' := 'call'}
PROPERTY PUBLIC ResetCount : UINT //! Recorded ResetCount for command-order verification.
GET
ResetCount := FResetCount;
END_GET
END_PROPERTY

{region 'Documentation'}
(*!
<summary>Recorded ResetOrder for command-order verification.</summary>
*)
{endregion}
{attribute 'monitoring' := 'call'}
PROPERTY PUBLIC ResetOrder : UINT //! Recorded ResetOrder for command-order verification.
GET
ResetOrder := FResetOrder;
END_GET
END_PROPERTY

END_FUNCTION_BLOCK

// ---- SelfTests/TestCases/TestSuite_EventBufferReset/Helper/BufferResetRunControlProbe.TcPOU
{region 'Documentation'}
(*!
<summary>Run Control using two borrowed Suite doubles and the existing controlled Orchestrator.</summary>
<description>
Bind and BindChildren precede Initialize. The real base handles external Buffer commands and
lifecycle; only scheduling is controlled so an Idle Orchestrator cannot add unrelated release calls.
ProcessTestSuites calls both borrowed concrete children once and presents stable Idle observations.
References remain valid for the enclosing Test Case lifetime. No production buffer command is replaced.
</description>
*)
{endregion}
FUNCTION_BLOCK BufferResetRunControlProbe EXTENDS RunControlBase
VAR
    FFirstSuite : REFERENCE TO BufferReleaseSuiteDouble;
    FSecondSuite : REFERENCE TO BufferReleaseSuiteDouble;
    FSuites : ARRAY[4..5] OF I_TestSuite;
    FIdleObservation : ST_OrchestrationObservation;
END_VAR

SUPER^(ControlData := ControlData);

{region 'Documentation'}
(*!
<summary>Selects isolated dependencies before production Initialize.</summary>
*)
{endregion}
METHOD PUBLIC Bind
VAR_INPUT
    Publisher : I_EventPublisher; //! Nonzero isolated event publisher retained before subject initialization; keep it alive through all subject use.
    Helper : I_Orchestrator; //! Nonzero injected orchestration helper retained before owner initialization; keep it alive through subject use.
END_VAR
FEventPublisher := Publisher;
FOrchestrator := Helper;
END_METHOD

{region 'Documentation'}
(*!
<summary>Binds the test-owned concrete Suites before root initialization.</summary>
*)
{endregion}
METHOD PUBLIC BindChildren
VAR_IN_OUT
    {attribute 'analysis' := '-167'}
    FirstSuite : BufferReleaseSuiteDouble; //! First borrowed Suite double retained by reference; keep it alive through subject use.
    {attribute 'analysis' := '-167'}
    SecondSuite : BufferReleaseSuiteDouble; //! Second borrowed Suite double retained by reference; keep it alive through subject use.
END_VAR
FFirstSuite REF= FirstSuite;
FSecondSuite REF= SecondSuite;
END_METHOD

{region 'Documentation'}
(*!
<summary>Registers both controlled Suites in stable order.</summary>
*)
{endregion}
METHOD PROTECTED Configure
VAR_IN_OUT
    // SA0167: Borrowed setup builder.
    {attribute 'analysis' := '-167'}
    Builder : RunControlConfigurationBuilder; //! Borrowed owner configuration builder used only during this Configure call; register this owner's concrete children.
END_VAR
FIdleObservation.State := E_State.Idle;
FIdleObservation.Result := E_Result.NotEvaluated;
FIdleObservation.Ready := TRUE;
FIdleObservation.Complete := FALSE;
FFirstSuite.Initialize(Name := CONCAT(Name, '.First'),
    Slot := 0);
FSecondSuite.Initialize(Name := CONCAT(Name, '.Second'),
    Slot := 0);
Builder.Initialize(Mode := E_OrchestrationMode.Serial,
    TestSuites := FSuites);
Builder.Register(TestSuite := FFirstSuite);
Builder.Register(TestSuite := FSecondSuite);
END_METHOD

{region 'Documentation'}
(*!
<summary>Returns the concrete registered Suite at its actual array index.</summary>
*)
{endregion}
METHOD PUBLIC GetTestSuite : I_TestSuite //! Typed Suite interface at the original array index; zero when no entry is available.
VAR_INPUT
    Index : DINT; //! Original occupied child-array index, rather than an ordinal position.
END_VAR
GetTestSuite := 0;
IF (Index < LOWER_BOUND(FSuites, 1)) OR (Index > UPPER_BOUND(FSuites, 1)) THEN
    RETURN;
END_IF;
GetTestSuite := FSuites[Index];
END_METHOD

{region 'Documentation'}
(*!
<summary>Calls both controlled children once; does not perform reservation work.</summary>
*)
{endregion}
METHOD PROTECTED ProcessTestSuites
FFirstSuite(ObservationInput := FIdleObservation);
FSecondSuite(ObservationInput := FIdleObservation);
END_METHOD

END_FUNCTION_BLOCK

// ---- SelfTests/TestCases/TestSuite_EventBufferReset/Helper/BufferReleaseSuiteDouble.TcPOU
{region 'Documentation'}
(*!
<summary>Controlled Suite release boundary with a real local buffer contribution.</summary>
<description>
PrepareRelease borrows the test-owned buffer and reserves a fixed contribution through its public API.
A rejected release deliberately retains that contribution. Later hard reset clears only the buffer
aggregate, not this failed local value. This double does not simulate a child hierarchy or admission
policy; the real hierarchy is exercised separately. No production state is modified for fault injection.
</description>
*)
{endregion}
FUNCTION_BLOCK BufferReleaseSuiteDouble EXTENDS RunControlSuiteDouble
VAR
    FBuffer : REFERENCE TO BufferCommandProbe;
    FContribution : UINT;
    FRejectRelease : BOOL;
    FReleaseOrder : UINT;
    FReleaseCount : UINT;
END_VAR

SUPER^(ObservationInput := ObservationInput);

{region 'Documentation'}
(*!
<summary>Records every attempt; selected failure retains the local contribution.</summary>
*)
{endregion}
METHOD PUBLIC FreeReservedEvents : BOOL //! TRUE when the contribution was released; FALSE for scripted rejection or inherited buffer release failure.
FReleaseCount := FReleaseCount + 1;
FReleaseOrder := FBuffer.RecordRelease();
FreeReservedEvents := FALSE;
IF FRejectRelease THEN
    RETURN;
END_IF;
FreeReservedEvents := FBuffer.FreeReservedSpace(EntryCount := FContribution,
    OwnerReservedEntryCount := FContribution);
END_METHOD

{region 'Documentation'}
(*!
<summary>Binds stable local storage and reserves the controlled Suite contribution.</summary>
*)
{endregion}
METHOD PUBLIC PrepareRelease : BOOL //! TRUE when the requested test contribution was reserved in the borrowed buffer.
VAR_INPUT
    RejectRelease : BOOL; //! TRUE makes subsequent release calls reject without freeing the contribution.
    EntryCount : UINT; //! Number of entries requested for this Suite double with zero headroom.
END_VAR
VAR_IN_OUT
    // SA0167: Borrowed test-owned buffer; no temporary instance.
    {attribute 'analysis' := '-167'}
    Buffer : BufferCommandProbe; //! Borrowed test-owned buffer retained for reservation and release; keep it alive until the binding is replaced.
END_VAR
FBuffer REF= Buffer;
FContribution := 0;
FRejectRelease := RejectRelease;
FReleaseOrder := 0;
FReleaseCount := 0;
PrepareRelease := FBuffer.ReserveSpace(EntryCount := EntryCount,
    HeadroomEntryCount := 0,
    OwnerReservedEntryCount := FContribution);
END_METHOD

{region 'Documentation'}
(*!
<summary>Recorded ReleaseCount for command-order verification.</summary>
*)
{endregion}
{attribute 'monitoring' := 'call'}
PROPERTY PUBLIC ReleaseCount : UINT //! Recorded ReleaseCount for command-order verification.
GET
ReleaseCount := FReleaseCount;
END_GET
END_PROPERTY

{region 'Documentation'}
(*!
<summary>Recorded ReleaseOrder for command-order verification.</summary>
*)
{endregion}
{attribute 'monitoring' := 'call'}
PROPERTY PUBLIC ReleaseOrder : UINT //! Recorded ReleaseOrder for command-order verification.
GET
ReleaseOrder := FReleaseOrder;
END_GET
END_PROPERTY

{region 'Documentation'}
(*!
<summary>Recorded ReservedEntryCount for command-order verification.</summary>
*)
{endregion}
{attribute 'monitoring' := 'call'}
PROPERTY PUBLIC ReservedEntryCount : UINT //! Recorded ReservedEntryCount for command-order verification.
GET
ReservedEntryCount := FContribution;
END_GET
END_PROPERTY

END_FUNCTION_BLOCK

// ---- SelfTests/TestCases/TestSuite_EventBufferReset/Test_BufferResetActiveRun.TcPOU
{region 'Documentation'}
(*!
<summary>Checks a hard Buffer Reset during a real reserved run and its normal orchestration error path.</summary>
<description>
The existing real root, Suite and Test Cases are called once per test cycle with isolated event storage.
Reset is submitted only after the first child is Running with a reservation. A thin buffer probe
captures the reset boundary before normal lifecycle processing can refill the new epoch.
Error-driven Abort afterwards is expected; no additional lifecycle Reset or automatic restart is requested.
New-epoch event checks retain all events until completion and reject loss or capacity exhaustion.
The real subject binds only local storage; expected findings remain in that storage.
Checking Assertions retain the outer selftest publisher. Each run reinitializes the subject.
</description>
*)
{endregion}
FUNCTION_BLOCK Test_BufferResetActiveRun EXTENDS TestCaseBase
VAR
    FSubject : ActiveResetBufferProbe;
    FEvents : ARRAY[1..BufferLength] OF ST_Event;
    FFifo : ST_FifoStatus;
    FBufferStatus : ST_EventBufferStatus;
    FPerformed : BOOL;
    FChecked : BOOL;
    FRoot : RunControlIntegrationSubject;
    FControl : ST_RunControl;
    FSuite : I_TestSuite;
    FChild : I_TestCase;
    FSecondChild : I_TestCase;
    FPhase : USINT;
    FActiveRun : AssertTrue;
    FActiveRunMatches : BOOL;
    FResetBoundary : AssertTrue;
    FResetBoundaryMatches : BOOL;
    FReservationsReleased : AssertTrue;
    FReservationsReleasedMatches : BOOL;
    FErrorPath : AssertTrue;
    FErrorPathMatches : BOOL;
    FNoLifecycleReset : AssertTrue;
    FNoLifecycleResetMatches : BOOL;
    FNewEpoch : AssertTrue;
    FNewEpochMatches : BOOL;
    FFinalization : AssertTrue;
    FFinalizationMatches : BOOL;
    FConfigurationPreserved : AssertTrue;
    FConfigurationPreservedMatches : BOOL;
END_VAR
VAR CONSTANT
    BufferLength : UINT := 257;
    SetupPhase : USINT := 0;
    AwaitIdlePhase : USINT := 1;
    AwaitActivePhase : USINT := 2;
    ResetPhase : USINT := 3;
    AwaitCompletionPhase : USINT := 4;
    OldEpochMarker : STRING := 'Discarded active-run marker';
END_VAR

SUPER^();

{region 'Documentation'}
(*!
<summary>Contributes each checking Assertion once.</summary>
*)
{endregion}
METHOD PROTECTED AggregateResults
VAR_INPUT
    Aggregator : I_ResultAggregator; //! Borrowed result sink owned by the outer Test Case; add this test's checking Assertions without resetting or retaining the sink.
END_VAR
Aggregator.AddProvider(Provider := FActiveRun);
Aggregator.AddProvider(Provider := FResetBoundary);
Aggregator.AddProvider(Provider := FReservationsReleased);
Aggregator.AddProvider(Provider := FErrorPath);
Aggregator.AddProvider(Provider := FNoLifecycleReset);
Aggregator.AddProvider(Provider := FNewEpoch);
Aggregator.AddProvider(Provider := FFinalization);
Aggregator.AddProvider(Provider := FConfigurationPreserved);
END_METHOD

{region 'Documentation'}
(*!
<summary>Requires all checking Assertions to be initialized.</summary>
*)
{endregion}
METHOD PROTECTED CheckInitialization : BOOL //! TRUE when the inherited initialization check and this concrete fixture check both accept the setup.
CheckInitialization := FALSE;
IF NOT SUPER^.CheckInitialization() THEN
    RETURN;
END_IF;

CheckInitialization := FActiveRun.IsInitialized
    AND FResetBoundary.IsInitialized
    AND FReservationsReleased.IsInitialized
    AND FErrorPath.IsInitialized
    AND FNoLifecycleReset.IsInitialized
    AND FNewEpoch.IsInitialized
    AND FFinalization.IsInitialized
    AND FConfigurationPreserved.IsInitialized;
END_METHOD

{region 'Documentation'}
(*!
<summary>Checks the retained new epoch for the existing error path and stable root finalization.</summary>
*)
{endregion}
METHOD PRIVATE CheckNewEpoch
VAR
    Index : UINT;
    MissingReservationReported : BOOL;
    RootErrorResultCount : UINT;
    RootCompletedCount : UINT;
END_VAR
FNewEpochMatches := (FFifo.ElementCount > 0) AND (FFifo.ElementCount < BufferLength - 1)
    AND (FFifo.IndexOut = 1) AND NOT FFifo.BufferFull AND NOT FFifo.BufferAlmostFull
    AND (FBufferStatus.LostEventCount = 0) AND (FBufferStatus.DeletedSequenceId = 0)
    AND (FBufferStatus.SequenceId = UINT_TO_UDINT(FFifo.ElementCount));
FNoLifecycleResetMatches := TRUE;
FOR Index := 1 TO FFifo.ElementCount DO
    FNewEpochMatches := FNewEpochMatches AND (FEvents[Index].SequenceId = UINT_TO_UDINT(Index))
        AND (FEvents[Index].Message <> OldEpochMarker);
    IF (FEvents[Index].EventType = E_EventType.Framework)
        AND (FEvents[Index].Severity = E_EventSeverity.Error)
        AND ((FEvents[Index].Message = CONCAT('Active child has no event reservation: ', FSuite.Name))
            OR (FEvents[Index].Message = CONCAT('Active child has no event reservation: ', FChild.Name))) THEN
        MissingReservationReported := TRUE;
    END_IF;
    IF (FEvents[Index].EventType = E_EventType.StateTransition)
        AND (FEvents[Index].State = E_State.Reset) THEN
        FNoLifecycleResetMatches := FALSE;
    END_IF;
    IF (FEvents[Index].Name = FRoot.Name) AND (FEvents[Index].OwnerScope = E_OwnerScope.RunControl) THEN
        IF (FEvents[Index].EventType = E_EventType.Result)
            AND (FEvents[Index].Result = E_Result.Error) THEN
            RootErrorResultCount := RootErrorResultCount + 1;
        END_IF;
        IF (FEvents[Index].EventType = E_EventType.StateTransition)
            AND (FEvents[Index].State = E_State.Completed) THEN
            RootCompletedCount := RootCompletedCount + 1;
        END_IF;
    END_IF;
END_FOR;
FErrorPathMatches := MissingReservationReported;
FFinalizationMatches := (RootErrorResultCount = 1) AND (RootCompletedCount = 1);
END_METHOD

{region 'Documentation'}
(*!
<summary>Initializes the checking Assertions for one test state.</summary>
*)
{endregion}
METHOD PROTECTED Configure
FPreparationStateCount := 0;
FTestStateCount := 1;
FActiveRun.Initialize(Parent := THIS^,
    AssertionName := 'ActiveRun');
FResetBoundary.Initialize(Parent := THIS^,
    AssertionName := 'ResetBoundary');
FReservationsReleased.Initialize(Parent := THIS^,
    AssertionName := 'ReservationsReleased');
FErrorPath.Initialize(Parent := THIS^,
    AssertionName := 'ErrorPath');
FNoLifecycleReset.Initialize(Parent := THIS^,
    AssertionName := 'NoLifecycleReset');
FNewEpoch.Initialize(Parent := THIS^,
    AssertionName := 'NewEpoch');
FFinalization.Initialize(Parent := THIS^,
    AssertionName := 'Finalization');
FConfigurationPreserved.Initialize(Parent := THIS^,
    AssertionName := 'ConfigurationPreserved');
END_METHOD

{region 'Documentation'}
(*!
<summary>Completes abort without asynchronous work.</summary>
*)
{endregion}
METHOD PROTECTED ProcessAbort
VAR_INPUT
    Enable : BOOL; //! Phase permission supplied by the owning Test Case; FALSE does not authorize progression, while observation may continue.
END_VAR
IF Enable THEN
    CompleteAbort();
END_IF;
END_METHOD

